screen "Screen_5" 800x480, template "Keep_1"
   Circle "Circle_2" at 38,164 size 32x32
      Appearance <- "Barcode181"
   Circle "Circle_1" at 38,224 size 32x32
      Appearance <- "Barcode190"
   Circle "Circle_3" at 38,279 size 32x32
      Appearance <- "Barcode199"
   Circle "Circle_4" at 38,336 size 32x32
      Appearance <- "Barcode208"
   Circle "Circle_5" at 38,393 size 32x32
      Appearance <- "Barcode217"
   Circle "Circle_6" at 102,164 size 32x32
      Appearance <- "Barcode182"
   Circle "Circle_7" at 102,224 size 32x32
      Appearance <- "Barcode191"
   Circle "Circle_8" at 102,279 size 32x32
      Appearance <- "Barcode200"
   Circle "Circle_9" at 102,336 size 32x32
      Appearance <- "Barcode209"
   Circle "Circle_10" at 102,393 size 32x32
      Appearance <- "Barcode218"
   Circle "Circle_11" at 166,164 size 32x32
      Appearance <- "Barcode183"
   Circle "Circle_12" at 166,224 size 32x32
      Appearance <- "Barcode192"
   Circle "Circle_13" at 166,279 size 32x32
      Appearance <- "Barcode201"
   Circle "Circle_14" at 166,336 size 32x32
      Appearance <- "Barcode210"
   Circle "Circle_15" at 166,393 size 32x32
      Appearance <- "Barcode219"
   Circle "Circle_16" at 230,164 size 32x32
      Appearance <- "Barcode184"
   Circle "Circle_17" at 230,224 size 32x32
      Appearance <- "Barcode193"
   Circle "Circle_18" at 230,279 size 32x32
      Appearance <- "Barcode202"
   Circle "Circle_19" at 230,336 size 32x32
      Appearance <- "Barcode211"
   Circle "Circle_20" at 230,393 size 32x32
      Appearance <- "Barcode220"
   Circle "Circle_21" at 294,164 size 32x32
      Appearance <- "Barcode185"
   Circle "Circle_22" at 294,224 size 32x32
      Appearance <- "Barcode194"
   Circle "Circle_23" at 294,279 size 32x32
      Appearance <- "Barcode203"
   Circle "Circle_24" at 294,336 size 32x32
      Appearance <- "Barcode212"
   Circle "Circle_25" at 294,393 size 32x32
      Appearance <- "Barcode221"
   Circle "Circle_26" at 358,164 size 32x32
      Appearance <- "Barcode186"
   Circle "Circle_27" at 358,225 size 32x32
      Appearance <- "Barcode195"
   Circle "Circle_28" at 358,279 size 32x32
      Appearance <- "Barcode204"
   Circle "Circle_29" at 358,336 size 32x32
      Appearance <- "Barcode213"
   Circle "Circle_30" at 358,393 size 32x32
      Appearance <- "Barcode222"
   Circle "Circle_31" at 422,164 size 32x32
      Appearance <- "Barcode187"
   Circle "Circle_32" at 422,224 size 32x32
      Appearance <- "Barcode196"
   Circle "Circle_33" at 422,279 size 32x32
      Appearance <- "Barcode205"
   Circle "Circle_34" at 422,336 size 32x32
      Appearance <- "Barcode214"
   Circle "Circle_35" at 422,393 size 32x32
      Appearance <- "Barcode223"
   Circle "Circle_36" at 486,164 size 32x32
      Appearance <- "Barcode188"
   Circle "Circle_37" at 486,224 size 32x32
      Appearance <- "Barcode197"
   Circle "Circle_38" at 486,279 size 32x32
      Appearance <- "Barcode206"
   Circle "Circle_39" at 486,336 size 32x32
      Appearance <- "Barcode215"
   Circle "Circle_40" at 486,393 size 32x32
      Appearance <- "Barcode224"
   Circle "Circle_41" at 550,163 size 32x32
      Appearance <- "Barcode189"
   Circle "Circle_42" at 550,224 size 32x32
      Appearance <- "Barcode198"
   Circle "Circle_43" at 550,279 size 32x32
      Appearance <- "Barcode207"
   Circle "Circle_44" at 550,336 size 32x32
      Appearance <- "Barcode216"
   Circle "Circle_45" at 550,393 size 32x32
      Appearance <- "Barcode225"
   TextField "Text field_8" at 473,145 size 66x20; Text 'Box_188'
   TextField "Text field_10" at 25,206 size 66x20; Text 'Box_190'
   TextField "Text field_11" at 88,206 size 66x20; Text 'Box_191'
   TextField "Text field_12" at 153,206 size 66x20; Text 'Box_192'
   TextField "Text field_13" at 217,206 size 66x20; Text 'Box_193'
   TextField "Text field_14" at 281,206 size 66x20; Text 'Box_194'
   TextField "Text field_15" at 345,206 size 66x20; Text 'Box_195'
   TextField "Text field_16" at 410,206 size 66x20; Text 'Box_196'
   TextField "Text field_17" at 473,206 size 66x20; Text 'Box_197'
   TextField "Text field_19" at 26,261 size 66x20; Text 'Box_199'
   TextField "Text field_20" at 89,261 size 66x20; Text 'Box_200'
   TextField "Text field_21" at 153,261 size 66x20; Text 'Box_201'
   TextField "Text field_22" at 217,261 size 66x20; Text 'Box_202'
   TextField "Text field_23" at 281,261 size 66x20; Text 'Box_203'
   TextField "Text field_24" at 346,261 size 66x20; Text 'Box_204'
   TextField "Text field_25" at 409,261 size 66x20; Text 'Box_205'
   TextField "Text field_26" at 473,261 size 66x20; Text 'Box_206'
   TextField "Text field_28" at 25,317 size 66x20; Text 'Box_208'
   TextField "Text field_29" at 88,317 size 66x20; Text 'Box_209'
   TextField "Text field_30" at 153,317 size 66x20; Text 'Box_210'
   TextField "Text field_31" at 218,317 size 66x20; Text 'Box_211'
   TextField "Text field_32" at 282,317 size 66x20; Text 'Box_212'
   TextField "Text field_33" at 346,317 size 66x20; Text 'Box_213'
   TextField "Text field_34" at 410,317 size 66x20; Text 'Box_214'
   TextField "Text field_35" at 472,317 size 66x20; Text 'Box_215'
   TextField "Text field_37" at 26,375 size 66x20; Text 'Box_217'
   TextField "Text field_38" at 88,375 size 66x20; Text 'Box_218'
   TextField "Text field_39" at 153,375 size 66x20; Text 'Box_219'
   TextField "Text field_40" at 217,375 size 66x20; Text 'Box_220'
   TextField "Text field_41" at 281,375 size 66x20; Text 'Box_221'
   TextField "Text field_42" at 345,375 size 66x20; Text 'Box_222'
   TextField "Text field_43" at 409,375 size 66x20; Text 'Box_223'
   TextField "Text field_44" at 473,375 size 66x20; Text 'Box_224'
   TextField "Text field_1" at 24,145 size 66x20; Text 'Box_181'
   TextField "Text field_2" at 87,145 size 66x20; Text 'Box_182'
   TextField "Text field_3" at 152,145 size 66x20; Text 'Box_183'
   TextField "Text field_4" at 216,145 size 66x20; Text 'Box_184'
   TextField "Text field_5" at 280,145 size 66x20; Text 'Box_185'
   TextField "Text field_6" at 344,145 size 66x20; Text 'Box_186'
   TextField "Text field_7" at 409,145 size 66x20; Text 'Box_187'
   TextField "Text field_9" at 536,145 size 66x20; Text 'Box_189'
   TextField "Text field_18" at 537,206 size 66x20; Text 'Box_198'
   TextField "Text field_27" at 537,261 size 66x20; Text 'Box_207'
   TextField "Text field_36" at 537,317 size 66x20; Text 'Box_216'
   TextField "Text field_45" at 536,375 size 66x20; Text 'Box_225'
   SymbolicIOField "Symbolic I/O field_1" at 621,342 size 167x24; TextOn '1'; TextOff '0'; TextList "BOX_All"
      ProcessValue <- "แสดงชื่อยา2"
   IOField "I/O field_1" at 624,160 size 160x64; FormatPattern ???????????
      on OnFinishInput: "Test2"(); "Storage"()
      ProcessValue <- "Expected/Value_All_V"
   TextField "Text field_47" at 648,418 size 78x17; Text ': Low Stock'
   TextField "Text field_46" at 646,395 size 104x17; Text ': Medium Stock'
   TextField "Text field_48" at 646,372 size 82x17; Text ': High Stock'
   GraphicView "Template_Graphic view_6" at 16,8 size 70x68; Picture "KMUTNB-Photoroom"
   GraphicView "Template_Graphic view_5" at 657,59 size 104x124; Picture "channels4_profile-Photoroom"
   Button "Button_5" at 633,292 size 64x24; TextOff 'Back'
      on Click: ActivateScreen("Screen_4", 0)
   Button "Button_6" at 716,292 size 64x24; TextOff 'Next'
      on Click: ActivateScreen("Screen_6", 0)
   GraphicView "Template_Graphic view_1" at 736,255 size 28x26; Picture "NEW_HOME"
   GraphicView "Template_Graphic view_2" at 650,253 size 28x27; Picture "play"
   GraphicView "Template_Graphic view_3" at 721,296 size 20x17; Picture "next-track"
   GraphicView "Template_Graphic view_4" at 638,296 size 20x17; Picture "previous-track"
   Button "Button_3" at 707,246 size 80x42; TextOn 'LOGOUT'; TextOff 'Text'
      on Activate: function_f23ef4c9(); ActivateScreen("1_OVERVIEW_1", 0)
   Button "Button_1" at 623,245 size 80x42; TextOff 'Text'
      on Press: SetTag("มีการปุ่มกดยืนยัน", 1)
      on Release: SetTag("มีการปุ่มกดยืนยัน", 0)
      on Activate: "Storage"()
      on Click: "Conveyor"(); ActivateScreen("Status System", 0)
   TextField "Text field_49" at 734,229 size 32x14; Text 'HOME'
   TextField "Text field_50" at 625,229 size 95x16; Text 'Simmulation Conveyor'

screen "Screen_6" 800x480, template "Keep_1"
   Circle "Circle_2" at 38,164 size 32x32
      Appearance <- "Barcode226"
   Circle "Circle_1" at 38,224 size 32x32
      Appearance <- "Barcode235"
   Circle "Circle_3" at 38,279 size 32x32
      Appearance <- "Barcode244"
   Circle "Circle_4" at 38,336 size 32x32
      Appearance <- "Barcode253"
   Circle "Circle_5" at 38,393 size 32x32
      Appearance <- "Barcode262"
   Circle "Circle_6" at 102,164 size 32x32
      Appearance <- "Barcode227"
   Circle "Circle_7" at 102,224 size 32x32
      Appearance <- "Barcode236"
   Circle "Circle_8" at 102,279 size 32x32
      Appearance <- "Barcode245"
   Circle "Circle_9" at 102,336 size 32x32
      Appearance <- "Barcode254"
   Circle "Circle_10" at 102,393 size 32x32
      Appearance <- "Barcode263"
   Circle "Circle_11" at 166,164 size 32x32
      Appearance <- "Barcode228"
   Circle "Circle_12" at 166,224 size 32x32
      Appearance <- "Barcode237"
   Circle "Circle_13" at 166,279 size 32x32
      Appearance <- "Barcode246"
   Circle "Circle_14" at 166,336 size 32x32
      Appearance <- "Barcode255"
   Circle "Circle_15" at 166,393 size 32x32
      Appearance <- "Barcode264"
   Circle "Circle_16" at 230,164 size 32x32
      Appearance <- "Barcode229"
   Circle "Circle_17" at 230,224 size 32x32
      Appearance <- "Barcode238"
   Circle "Circle_18" at 230,279 size 32x32
      Appearance <- "Barcode247"
   Circle "Circle_19" at 230,336 size 32x32
      Appearance <- "Barcode256"
   Circle "Circle_20" at 230,393 size 32x32
      Appearance <- "Barcode265"
   Circle "Circle_21" at 294,164 size 32x32
      Appearance <- "Barcode230"
   Circle "Circle_22" at 294,224 size 32x32
      Appearance <- "Barcode239"
   Circle "Circle_23" at 294,279 size 32x32
      Appearance <- "Barcode248"
   Circle "Circle_24" at 294,336 size 32x32
      Appearance <- "Barcode257"
   Circle "Circle_25" at 294,393 size 32x32
      Appearance <- "Barcode266"
   Circle "Circle_26" at 358,164 size 32x32
      Appearance <- "Barcode231"
   Circle "Circle_27" at 358,225 size 32x32
      Appearance <- "Barcode240"
   Circle "Circle_28" at 358,279 size 32x32
      Appearance <- "Barcode249"
   Circle "Circle_29" at 358,336 size 32x32
      Appearance <- "Barcode258"
   Circle "Circle_30" at 358,393 size 32x32
      Appearance <- "Barcode267"
   Circle "Circle_31" at 422,164 size 32x32
      Appearance <- "Barcode232"
   Circle "Circle_32" at 422,224 size 32x32
      Appearance <- "Barcode241"
   Circle "Circle_33" at 422,279 size 32x32
      Appearance <- "Barcode250"
   Circle "Circle_34" at 422,336 size 32x32
      Appearance <- "Barcode259"
   Circle "Circle_35" at 422,393 size 32x32
      Appearance <- "Barcode268"
   Circle "Circle_36" at 486,164 size 32x32
      Appearance <- "Barcode233"
   Circle "Circle_37" at 486,224 size 32x32
      Appearance <- "Barcode242"
   Circle "Circle_38" at 486,279 size 32x32
      Appearance <- "Barcode251"
   Circle "Circle_39" at 486,336 size 32x32
      Appearance <- "Barcode260"
   Circle "Circle_40" at 486,393 size 32x32
      Appearance <- "Barcode269"
   Circle "Circle_41" at 550,163 size 32x32
      Appearance <- "Barcode234"
   Circle "Circle_42" at 550,224 size 32x32
      Appearance <- "Barcode243"
   Circle "Circle_43" at 550,279 size 32x32
      Appearance <- "Barcode252"
   Circle "Circle_44" at 550,336 size 32x32
      Appearance <- "Barcode261"
   Circle "Circle_45" at 550,393 size 32x32
      Appearance <- "Barcode270"
   TextField "Text field_8" at 473,145 size 66x20; Text 'Box_233'
   TextField "Text field_10" at 25,206 size 66x20; Text 'Box_235'
   TextField "Text field_11" at 88,206 size 66x20; Text 'Box_236'
   TextField "Text field_12" at 153,206 size 66x20; Text 'Box_237'
   TextField "Text field_13" at 217,206 size 66x20; Text 'Box_238'
   TextField "Text field_14" at 281,206 size 66x20; Text 'Box_239'
   TextField "Text field_15" at 345,206 size 66x20; Text 'Box_240'
   TextField "Text field_16" at 410,206 size 66x20; Text 'Box_241'
   TextField "Text field_17" at 473,206 size 66x20; Text 'Box_242'
   TextField "Text field_19" at 26,261 size 66x20; Text 'Box_244'
   TextField "Text field_20" at 89,261 size 66x20; Text 'Box_245'
   TextField "Text field_21" at 153,261 size 66x20; Text 'Box_246'
   TextField "Text field_22" at 217,261 size 66x20; Text 'Box_247'
   TextField "Text field_23" at 281,261 size 66x20; Text 'Box_248'
   TextField "Text field_24" at 346,261 size 66x20; Text 'Box_249'
   TextField "Text field_25" at 409,261 size 66x20; Text 'Box_250'
   TextField "Text field_26" at 473,261 size 66x20; Text 'Box_251'
   TextField "Text field_28" at 25,317 size 66x20; Text 'Box_253'
   TextField "Text field_29" at 88,317 size 66x20; Text 'Box_254'
   TextField "Text field_30" at 153,317 size 66x20; Text 'Box_255'
   TextField "Text field_31" at 217,317 size 66x20; Text 'Box_256'
   TextField "Text field_32" at 281,317 size 66x20; Text 'Box_257'
   TextField "Text field_33" at 344,317 size 66x20; Text 'Box_258'
   TextField "Text field_34" at 409,317 size 66x20; Text 'Box_259'
   TextField "Text field_35" at 472,317 size 66x20; Text 'Box_260'
   TextField "Text field_37" at 24,375 size 66x20; Text 'Box_262'
   TextField "Text field_38" at 88,375 size 66x20; Text 'Box_263'
   TextField "Text field_39" at 153,375 size 66x20; Text 'Box_264'
   TextField "Text field_40" at 217,375 size 66x20; Text 'Box_265'
   TextField "Text field_41" at 281,375 size 66x20; Text 'Box_266'
   TextField "Text field_42" at 345,375 size 66x20; Text 'Box_267'
   TextField "Text field_43" at 409,375 size 66x20; Text 'Box_268'
   TextField "Text field_44" at 473,375 size 66x20; Text 'Box_269'
   TextField "Text field_1" at 24,145 size 66x20; Text 'Box_226'
   TextField "Text field_2" at 87,145 size 66x20; Text 'Box_227'
   TextField "Text field_3" at 152,145 size 66x20; Text 'Box_228'
   TextField "Text field_4" at 216,145 size 66x20; Text 'Box_229'
   TextField "Text field_5" at 280,145 size 66x20; Text 'Box_230'
   TextField "Text field_6" at 344,145 size 66x20; Text 'Box_231'
   TextField "Text field_7" at 409,145 size 66x20; Text 'Box_232'
   TextField "Text field_9" at 536,145 size 66x20; Text 'Box_234'
   TextField "Text field_18" at 537,206 size 66x20; Text 'Box_243'
   TextField "Text field_27" at 537,261 size 66x20; Text 'Box_252'
   TextField "Text field_36" at 537,317 size 66x20; Text 'Box_261'
   TextField "Text field_45" at 536,375 size 66x20; Text 'Box_270'
   SymbolicIOField "Symbolic I/O field_1" at 621,342 size 167x24; TextOn '1'; TextOff '0'; TextList "BOX_All"
      ProcessValue <- "แสดงชื่อยา2"
   IOField "I/O field_1" at 624,160 size 160x64; FormatPattern ???????????
      on OnFinishInput: "Test2"(); "Storage"()
      ProcessValue <- "Expected/Value_All_V"
   TextField "Text field_47" at 648,418 size 78x17; Text ': Low Stock'
   TextField "Text field_46" at 646,395 size 104x17; Text ': Medium Stock'
   TextField "Text field_48" at 646,372 size 82x17; Text ': High Stock'
   GraphicView "Template_Graphic view_6" at 16,8 size 70x68; Picture "KMUTNB-Photoroom"
   GraphicView "Template_Graphic view_5" at 657,59 size 104x124; Picture "channels4_profile-Photoroom"
   Button "Button_5" at 633,292 size 64x24; TextOff 'Back'
      on Click: ActivateScreen("Screen_5", 0)
   Button "Button_6" at 716,292 size 64x24; TextOff 'Next'
      on Click: ActivateScreen("Screen_7", 0)
   GraphicView "Template_Graphic view_1" at 736,255 size 28x26; Picture "NEW_HOME"
   GraphicView "Template_Graphic view_2" at 650,253 size 28x27; Picture "play"
   GraphicView "Template_Graphic view_3" at 721,296 size 20x17; Picture "next-track"
   GraphicView "Template_Graphic view_4" at 638,296 size 20x17; Picture "previous-track"
   Button "Button_3" at 707,246 size 80x42; TextOn 'LOGOUT'; TextOff 'Text'
      on Activate: function_f23ef4c9(); ActivateScreen("1_OVERVIEW_1", 0)
   Button "Button_1" at 623,245 size 80x42; TextOff 'Text'
      on Press: SetTag("มีการปุ่มกดยืนยัน", 1)
      on Release: SetTag("มีการปุ่มกดยืนยัน", 0)
      on Activate: "Storage"()
      on Click: "Conveyor"(); ActivateScreen("Status System", 0)
   TextField "Text field_49" at 734,229 size 32x14; Text 'HOME'
   TextField "Text field_50" at 625,229 size 95x16; Text 'Simmulation Conveyor'

screen "Screen_7" 800x480, template "Keep_1"
   Circle "Circle_2" at 38,164 size 32x32
      Appearance <- "Barcode271"
   Circle "Circle_1" at 38,224 size 32x32
      Appearance <- "Barcode280"
   Circle "Circle_3" at 38,279 size 32x32
      Appearance <- "Barcode289"
   Circle "Circle_4" at 38,336 size 32x32
      Appearance <- "Barcode298"
   Circle "Circle_5" at 38,393 size 32x32
      Appearance <- "Barcode307"
   Circle "Circle_6" at 102,164 size 32x32
      Appearance <- "Barcode272"
   Circle "Circle_7" at 102,224 size 32x32
      Appearance <- "Barcode281"
   Circle "Circle_8" at 102,279 size 32x32
      Appearance <- "Barcode290"
   Circle "Circle_9" at 102,336 size 32x32
      Appearance <- "Barcode299"
   Circle "Circle_10" at 102,393 size 32x32
      Appearance <- "Barcode308"
   Circle "Circle_11" at 166,164 size 32x32
      Appearance <- "Barcode273"
   Circle "Circle_12" at 166,224 size 32x32
      Appearance <- "Barcode282"
   Circle "Circle_13" at 166,279 size 32x32
      Appearance <- "Barcode291"
   Circle "Circle_14" at 166,336 size 32x32
      Appearance <- "Barcode300"
   Circle "Circle_15" at 166,393 size 32x32
      Appearance <- "Barcode309"
   Circle "Circle_16" at 230,164 size 32x32
      Appearance <- "Barcode274"
   Circle "Circle_17" at 230,224 size 32x32
      Appearance <- "Barcode283"
   Circle "Circle_18" at 230,279 size 32x32
      Appearance <- "Barcode292"
   Circle "Circle_19" at 230,336 size 32x32
      Appearance <- "Barcode301"
   Circle "Circle_20" at 230,393 size 32x32
      Appearance <- "Barcode310"
   Circle "Circle_21" at 294,164 size 32x32
      Appearance <- "Barcode275"
   Circle "Circle_22" at 294,224 size 32x32
      Appearance <- "Barcode284"
   Circle "Circle_23" at 294,279 size 32x32
      Appearance <- "Barcode293"
   Circle "Circle_24" at 294,336 size 32x32
      Appearance <- "Barcode302"
   Circle "Circle_25" at 294,393 size 32x32
      Appearance <- "Barcode311"
   Circle "Circle_26" at 358,164 size 32x32
      Appearance <- "Barcode276"
   Circle "Circle_27" at 358,225 size 32x32
      Appearance <- "Barcode285"
   Circle "Circle_28" at 358,279 size 32x32
      Appearance <- "Barcode294"
   Circle "Circle_29" at 358,336 size 32x32
      Appearance <- "Barcode303"
   Circle "Circle_30" at 358,393 size 32x32
      Appearance <- "Barcode312"
   Circle "Circle_31" at 422,164 size 32x32
      Appearance <- "Barcode277"
   Circle "Circle_32" at 422,224 size 32x32
      Appearance <- "Barcode286"
   Circle "Circle_33" at 422,279 size 32x32
      Appearance <- "Barcode295"
   Circle "Circle_34" at 422,336 size 32x32
      Appearance <- "Barcode304"
   Circle "Circle_35" at 422,393 size 32x32
      Appearance <- "Barcode313"
   Circle "Circle_36" at 486,164 size 32x32
      Appearance <- "Barcode278"
   Circle "Circle_37" at 486,224 size 32x32
      Appearance <- "Barcode287"
   Circle "Circle_38" at 486,279 size 32x32
      Appearance <- "Barcode296"
   Circle "Circle_39" at 486,336 size 32x32
      Appearance <- "Barcode305"
   Circle "Circle_40" at 486,393 size 32x32
      Appearance <- "Barcode314"
   Circle "Circle_41" at 550,163 size 32x32
      Appearance <- "Barcode279"
   Circle "Circle_42" at 550,224 size 32x32
      Appearance <- "Barcode288"
   Circle "Circle_43" at 550,279 size 32x32
      Appearance <- "Barcode297"
   Circle "Circle_44" at 550,336 size 32x32
      Appearance <- "Barcode306"
   Circle "Circle_45" at 550,393 size 32x32
      Appearance <- "Barcode315"
   TextField "Text field_8" at 473,145 size 66x20; Text 'Box_278'
   TextField "Text field_10" at 25,206 size 66x20; Text 'Box_280'
   TextField "Text field_11" at 88,206 size 66x20; Text 'Box_281'
   TextField "Text field_12" at 153,206 size 66x20; Text 'Box_282'
   TextField "Text field_13" at 217,206 size 66x20; Text 'Box_283'
   TextField "Text field_14" at 281,206 size 66x20; Text 'Box_284'
   TextField "Text field_15" at 345,206 size 66x20; Text 'Box_285'
   TextField "Text field_16" at 410,206 size 66x20; Text 'Box_286'
   TextField "Text field_17" at 473,206 size 66x20; Text 'Box_287'
   TextField "Text field_19" at 25,261 size 66x20; Text 'Box_289'
   TextField "Text field_20" at 89,261 size 66x20; Text 'Box_290'
   TextField "Text field_21" at 153,261 size 66x20; Text 'Box_291'
   TextField "Text field_22" at 217,261 size 66x20; Text 'Box_292'
   TextField "Text field_23" at 281,261 size 66x20; Text 'Box_293'
   TextField "Text field_24" at 346,261 size 66x20; Text 'Box_294'
   TextField "Text field_25" at 409,261 size 66x20; Text 'Box_295'
   TextField "Text field_26" at 473,261 size 66x20; Text 'Box_296'
   TextField "Text field_28" at 25,317 size 66x20; Text 'Box_298'
   TextField "Text field_29" at 88,317 size 66x20; Text 'Box_299'
   TextField "Text field_30" at 153,317 size 66x20; Text 'Box_300'
   TextField "Text field_31" at 217,317 size 66x20; Text 'Box_301'
   TextField "Text field_32" at 281,317 size 66x20; Text 'Box_302'
   TextField "Text field_33" at 344,317 size 66x20; Text 'Box_303'
   TextField "Text field_34" at 409,317 size 66x20; Text 'Box_304'
   TextField "Text field_35" at 472,317 size 66x20; Text 'Box_305'
   TextField "Text field_37" at 24,375 size 66x20; Text 'Box_307'
   TextField "Text field_38" at 88,375 size 66x20; Text 'Box_308'
   TextField "Text field_39" at 153,375 size 66x20; Text 'Box_309'
   TextField "Text field_40" at 217,375 size 66x20; Text 'Box_310'
   TextField "Text field_41" at 281,375 size 66x20; Text 'Box_311'
   TextField "Text field_42" at 345,375 size 66x20; Text 'Box_312'
   TextField "Text field_43" at 409,375 size 66x20; Text 'Box_313'
   TextField "Text field_44" at 473,375 size 66x20; Text 'Box_314'
   TextField "Text field_1" at 24,145 size 66x20; Text 'Box_271'
   TextField "Text field_2" at 87,145 size 66x20; Text 'Box_272'
   TextField "Text field_3" at 152,145 size 66x20; Text 'Box_273'
   TextField "Text field_4" at 216,145 size 66x20; Text 'Box_274'
   TextField "Text field_5" at 280,145 size 66x20; Text 'Box_275'
   TextField "Text field_6" at 344,145 size 66x20; Text 'Box_276'
   TextField "Text field_7" at 409,145 size 66x20; Text 'Box_277'
   TextField "Text field_9" at 536,145 size 66x20; Text 'Box_279'
   TextField "Text field_18" at 537,206 size 66x20; Text 'Box_288'
   TextField "Text field_27" at 537,261 size 66x20; Text 'Box_297'
   TextField "Text field_36" at 537,317 size 66x20; Text 'Box_306'
   TextField "Text field_45" at 536,375 size 66x20; Text 'Box_315'
   SymbolicIOField "Symbolic I/O field_1" at 621,342 size 167x24; TextOn '1'; TextOff '0'; TextList "BOX_All"
      ProcessValue <- "แสดงชื่อยา2"
   IOField "I/O field_1" at 624,160 size 160x64; FormatPattern ???????????
      on OnFinishInput: "Test2"(); "Storage"()
      ProcessValue <- "Expected/Value_All_V"
   TextField "Text field_47" at 648,418 size 78x17; Text ': Low Stock'
   TextField "Text field_46" at 646,395 size 104x17; Text ': Medium Stock'
   TextField "Text field_48" at 646,372 size 82x17; Text ': High Stock'
   GraphicView "Template_Graphic view_6" at 16,8 size 70x68; Picture "KMUTNB-Photoroom"
   GraphicView "Template_Graphic view_5" at 657,59 size 104x124; Picture "channels4_profile-Photoroom"
   Button "Button_5" at 633,292 size 64x24; TextOff 'Back'
      on Click: ActivateScreen("Screen_6", 0)
   Button "Button_6" at 716,292 size 64x24; TextOff 'Next'
      on Click: ActivateScreen("Screen_8", 0)
   GraphicView "Template_Graphic view_1" at 736,255 size 28x26; Picture "NEW_HOME"
   GraphicView "Template_Graphic view_2" at 650,253 size 28x27; Picture "play"
   GraphicView "Template_Graphic view_3" at 721,296 size 20x17; Picture "next-track"
   GraphicView "Template_Graphic view_4" at 638,296 size 20x17; Picture "previous-track"
   Button "Button_3" at 707,246 size 80x42; TextOn 'LOGOUT'; TextOff 'Text'
      on Activate: function_f23ef4c9(); ActivateScreen("1_OVERVIEW_1", 0)
   Button "Button_1" at 623,245 size 80x42; TextOff 'Text'
      on Press: SetTag("มีการปุ่มกดยืนยัน", 1)
      on Release: SetTag("มีการปุ่มกดยืนยัน", 0)
      on Activate: "Storage"()
      on Click: "Conveyor"(); ActivateScreen("Status System", 0)
   TextField "Text field_49" at 734,229 size 32x14; Text 'HOME'
   TextField "Text field_50" at 625,229 size 95x16; Text 'Simmulation Conveyor'

screen "Screen_8" 800x480, template "Keep_1"
   Circle "Circle_2" at 38,164 size 32x32
      Appearance <- "Barcode316"
   Circle "Circle_1" at 38,224 size 32x32
      Appearance <- "Barcode325"
   Circle "Circle_3" at 38,279 size 32x32
      Appearance <- "Barcode334"
   Circle "Circle_4" at 38,336 size 32x32
      Appearance <- "Barcode343"
   Circle "Circle_5" at 38,393 size 32x32
      Appearance <- "Barcode352"
   Circle "Circle_6" at 102,164 size 32x32
      Appearance <- "Barcode317"
   Circle "Circle_7" at 102,224 size 32x32
      Appearance <- "Barcode326"
   Circle "Circle_8" at 102,279 size 32x32
      Appearance <- "Barcode335"
   Circle "Circle_9" at 102,336 size 32x32
      Appearance <- "Barcode344"
   Circle "Circle_10" at 102,393 size 32x32
      Appearance <- "Barcode353"
   Circle "Circle_11" at 166,164 size 32x32
      Appearance <- "Barcode318"
   Circle "Circle_12" at 166,224 size 32x32
      Appearance <- "Barcode327"
   Circle "Circle_13" at 166,279 size 32x32
      Appearance <- "Barcode336"
   Circle "Circle_14" at 166,336 size 32x32
      Appearance <- "Barcode345"
   Circle "Circle_15" at 166,393 size 32x32
      Appearance <- "Barcode354"
   Circle "Circle_16" at 230,164 size 32x32
      Appearance <- "Barcode319"
   Circle "Circle_17" at 230,224 size 32x32
      Appearance <- "Barcode328"
   Circle "Circle_18" at 230,279 size 32x32
      Appearance <- "Barcode337"
   Circle "Circle_19" at 230,336 size 32x32
      Appearance <- "Barcode346"
   Circle "Circle_20" at 230,393 size 32x32
      Appearance <- "Barcode355"
   Circle "Circle_21" at 294,164 size 32x32
      Appearance <- "Barcode320"
   Circle "Circle_22" at 294,224 size 32x32
      Appearance <- "Barcode329"
   Circle "Circle_23" at 294,279 size 32x32
      Appearance <- "Barcode338"
   Circle "Circle_24" at 294,336 size 32x32
      Appearance <- "Barcode347"
   Circle "Circle_25" at 294,393 size 32x32
      Appearance <- "Barcode356"
   Circle "Circle_26" at 358,164 size 32x32
      Appearance <- "Barcode321"
   Circle "Circle_27" at 358,225 size 32x32
      Appearance <- "Barcode330"
   Circle "Circle_28" at 358,279 size 32x32
      Appearance <- "Barcode339"
   Circle "Circle_29" at 358,336 size 32x32
      Appearance <- "Barcode348"
   Circle "Circle_30" at 358,393 size 32x32
      Appearance <- "Barcode357"
   Circle "Circle_31" at 422,164 size 32x32
      Appearance <- "Barcode322"
   Circle "Circle_32" at 422,224 size 32x32
      Appearance <- "Barcode331"
   Circle "Circle_33" at 422,279 size 32x32
      Appearance <- "Barcode340"
   Circle "Circle_34" at 422,336 size 32x32
      Appearance <- "Barcode349"
   Circle "Circle_35" at 422,393 size 32x32
      Appearance <- "Barcode358"
   Circle "Circle_36" at 486,164 size 32x32
      Appearance <- "Barcode323"
   Circle "Circle_37" at 486,224 size 32x32
      Appearance <- "Barcode332"
   Circle "Circle_38" at 486,279 size 32x32
      Appearance <- "Barcode341"
   Circle "Circle_39" at 486,336 size 32x32
      Appearance <- "Barcode350"
   Circle "Circle_40" at 486,393 size 32x32
      Appearance <- "Barcode359"
   Circle "Circle_41" at 550,163 size 32x32
      Appearance <- "Barcode324"
   Circle "Circle_42" at 550,224 size 32x32
      Appearance <- "Barcode333"
   Circle "Circle_43" at 550,279 size 32x32
      Appearance <- "Barcode342"
   Circle "Circle_44" at 550,336 size 32x32
      Appearance <- "Barcode351"
   Circle "Circle_45" at 550,393 size 32x32
      Appearance <- "Barcode360"
   TextField "Text field_8" at 473,145 size 66x20; Text 'Box_323'
   TextField "Text field_10" at 25,206 size 66x20; Text 'Box_325'
   TextField "Text field_11" at 88,206 size 66x20; Text 'Box_326'
   TextField "Text field_12" at 153,206 size 66x20; Text 'Box_327'
   TextField "Text field_13" at 217,206 size 66x20; Text 'Box_328'
   TextField "Text field_14" at 281,206 size 66x20; Text 'Box_329'
   TextField "Text field_15" at 345,206 size 66x20; Text 'Box_330'
   TextField "Text field_16" at 410,206 size 66x20; Text 'Box_331'
   TextField "Text field_17" at 473,206 size 66x20; Text 'Box_332'
   TextField "Text field_19" at 25,261 size 66x20; Text 'Box_334'
   TextField "Text field_20" at 89,261 size 66x20; Text 'Box_335'
   TextField "Text field_21" at 153,261 size 66x20; Text 'Box_336'
   TextField "Text field_22" at 217,261 size 66x20; Text 'Box_337'
   TextField "Text field_23" at 281,261 size 66x20; Text 'Box_338'
   TextField "Text field_24" at 346,261 size 66x20; Text 'Box_339'
   TextField "Text field_25" at 409,261 size 66x20; Text 'Box_340'
   TextField "Text field_26" at 473,261 size 66x20; Text 'Box_341'
   TextField "Text field_28" at 25,317 size 66x20; Text 'Box_343'
   TextField "Text field_29" at 88,317 size 66x20; Text 'Box_344'
   TextField "Text field_30" at 153,317 size 66x20; Text 'Box_345'
   TextField "Text field_31" at 217,317 size 66x20; Text 'Box_346'
   TextField "Text field_32" at 281,317 size 66x20; Text 'Box_347'
   TextField "Text field_33" at 344,317 size 66x20; Text 'Box_348'
   TextField "Text field_34" at 409,317 size 66x20; Text 'Box_349'
   TextField "Text field_35" at 472,317 size 66x20; Text 'Box_350'
   TextField "Text field_37" at 24,375 size 66x20; Text 'Box_352'
   TextField "Text field_38" at 88,375 size 66x20; Text 'Box_353'
   TextField "Text field_39" at 153,375 size 66x20; Text 'Box_354'
   TextField "Text field_40" at 217,375 size 66x20; Text 'Box_355'
   TextField "Text field_41" at 281,375 size 66x20; Text 'Box_356'
   TextField "Text field_42" at 345,375 size 66x20; Text 'Box_357'
   TextField "Text field_43" at 409,375 size 66x20; Text 'Box_358'
   TextField "Text field_44" at 473,375 size 66x20; Text 'Box_359'
   TextField "Text field_1" at 24,145 size 66x20; Text 'Box_316'
   TextField "Text field_2" at 89,145 size 66x20; Text 'Box_317'
   TextField "Text field_3" at 152,145 size 66x20; Text 'Box_318'
   TextField "Text field_4" at 216,145 size 66x20; Text 'Box_319'
   TextField "Text field_5" at 280,145 size 66x20; Text 'Box_320'
   TextField "Text field_6" at 344,145 size 66x20; Text 'Box_321'
   TextField "Text field_7" at 409,145 size 66x20; Text 'Box_322'
   TextField "Text field_9" at 536,145 size 66x20; Text 'Box_324'
   TextField "Text field_18" at 537,206 size 66x20; Text 'Box_333'
   TextField "Text field_27" at 537,261 size 66x20; Text 'Box_342'
   TextField "Text field_36" at 537,317 size 66x20; Text 'Box_351'
   TextField "Text field_45" at 536,375 size 66x20; Text 'Box_360'
   SymbolicIOField "Symbolic I/O field_1" at 621,342 size 167x24; TextOn '1'; TextOff '0'; TextList "BOX_All"
      ProcessValue <- "แสดงชื่อยา2"
   IOField "I/O field_1" at 624,160 size 160x64; FormatPattern ???????????
      on OnFinishInput: "Test2"(); "Storage"()
      ProcessValue <- "Expected/Value_All_V"
   TextField "Text field_47" at 648,418 size 78x17; Text ': Low Stock'
   TextField "Text field_46" at 646,395 size 104x17; Text ': Medium Stock'
   TextField "Text field_48" at 646,372 size 82x17; Text ': High Stock'
   GraphicView "Template_Graphic view_6" at 16,8 size 70x68; Picture "KMUTNB-Photoroom"
   GraphicView "Template_Graphic view_5" at 657,59 size 104x124; Picture "channels4_profile-Photoroom"
   Button "Button_5" at 633,292 size 64x24; TextOff 'Back'
      on Click: ActivateScreen("Screen_7", 0)
   Button "Button_6" at 716,292 size 64x24; TextOff 'Next'
      on Click: ActivateScreen("Screen_9", 0)
   GraphicView "Template_Graphic view_1" at 736,255 size 28x26; Picture "NEW_HOME"
   GraphicView "Template_Graphic view_2" at 650,253 size 28x27; Picture "play"
   GraphicView "Template_Graphic view_3" at 721,296 size 20x17; Picture "next-track"
   GraphicView "Template_Graphic view_4" at 638,296 size 20x17; Picture "previous-track"
   Button "Button_3" at 707,246 size 80x42; TextOn 'LOGOUT'; TextOff 'Text'
      on Activate: function_f23ef4c9(); ActivateScreen("1_OVERVIEW_1", 0)
   Button "Button_1" at 623,245 size 80x42; TextOff 'Text'
      on Press: SetTag("มีการปุ่มกดยืนยัน", 1)
      on Release: SetTag("มีการปุ่มกดยืนยัน", 0)
      on Activate: "Storage"()
      on Click: "Conveyor"(); ActivateScreen("Status System", 0)
   TextField "Text field_49" at 734,229 size 32x14; Text 'HOME'
   TextField "Text field_50" at 625,229 size 95x16; Text 'Simmulation Conveyor'

screen "Screen_9" 800x480, template "Keep_1"
   TextField "Text field_8" at 473,145 size 66x20; Text 'Box_368'
   TextField "Text field_10" at 25,206 size 66x20; Text 'Box_370'
   TextField "Text field_11" at 88,206 size 66x20; Text 'Box_371'
   TextField "Text field_12" at 153,206 size 66x20; Text 'Box_372'
   TextField "Text field_13" at 217,206 size 66x20; Text 'Box_373'
   TextField "Text field_14" at 281,206 size 66x20; Text 'Box_374'
   TextField "Text field_15" at 345,206 size 66x20; Text 'Box_375'
   TextField "Text field_16" at 410,206 size 66x20; Text 'Box_376'
   TextField "Text field_17" at 473,206 size 66x20; Text 'Box_377'
   TextField "Text field_19" at 25,261 size 66x20; Text 'Box_379'
   TextField "Text field_20" at 89,261 size 66x20; Text 'Box_380'
   TextField "Text field_21" at 153,261 size 66x20; Text 'Box_381'
   TextField "Text field_22" at 217,261 size 66x20; Text 'Box_382'
   TextField "Text field_23" at 281,261 size 66x20; Text 'Box_383'
   TextField "Text field_24" at 346,261 size 66x20; Text 'Box_384'
   TextField "Text field_25" at 409,261 size 66x20; Text 'Box_385'
   TextField "Text field_26" at 473,261 size 66x20; Text 'Box_386'
   TextField "Text field_28" at 25,317 size 66x20; Text 'Box_388'
   TextField "Text field_29" at 88,317 size 66x20; Text 'Box_389'
   TextField "Text field_30" at 153,317 size 66x20; Text 'Box_390'
   TextField "Text field_31" at 217,317 size 66x20; Text 'Box_391'
   TextField "Text field_32" at 281,317 size 66x20; Text 'Box_392'
   TextField "Text field_33" at 344,317 size 66x20; Text 'Box_393'
   TextField "Text field_34" at 409,317 size 66x20; Text 'Box_394'
   TextField "Text field_35" at 472,317 size 66x20; Text 'Box_395'
   TextField "Text field_37" at 24,375 size 66x20; Text 'Box_397'
   TextField "Text field_38" at 88,375 size 66x20; Text 'Box_398'
   TextField "Text field_39" at 153,375 size 66x20; Text 'Box_399'
   TextField "Text field_40" at 217,375 size 66x20; Text 'Box_400'
   TextField "Text field_41" at 281,375 size 66x20; Text 'Box_401'
   TextField "Text field_42" at 345,375 size 66x20; Text 'Box_402'
   TextField "Text field_43" at 409,375 size 66x20; Text 'Box_403'
   TextField "Text field_44" at 473,375 size 66x20; Text 'Box_404'
   TextField "Text field_1" at 24,145 size 66x20; Text 'Box_361'
   TextField "Text field_2" at 89,145 size 66x20; Text 'Box_362'
   TextField "Text field_3" at 152,145 size 66x20; Text 'Box_363'
   TextField "Text field_4" at 216,145 size 66x20; Text 'Box_364'
   TextField "Text field_5" at 280,145 size 66x20; Text 'Box_365'
   TextField "Text field_6" at 344,145 size 66x20; Text 'Box_366'
   TextField "Text field_7" at 409,145 size 66x20; Text 'Box_367'
   TextField "Text field_9" at 536,145 size 66x20; Text 'Box_369'
   TextField "Text field_18" at 537,206 size 66x20; Text 'Box_378'
   TextField "Text field_27" at 537,261 size 66x20; Text 'Box_387'
   TextField "Text field_36" at 537,317 size 66x20; Text 'Box_396'
   TextField "Text field_45" at 536,375 size 66x20; Text 'Box_405'
   SymbolicIOField "Symbolic I/O field_1" at 621,342 size 167x24; TextOn '1'; TextOff '0'; TextList "BOX_All"
      ProcessValue <- "แสดงชื่อยา2"
   IOField "I/O field_1" at 624,160 size 160x64; FormatPattern ???????????
      on OnFinishInput: "Test2"(); "Storage"()
      ProcessValue <- "Expected/Value_All_V"
   TextField "Text field_47" at 648,418 size 78x17; Text ': Low Stock'
   TextField "Text field_46" at 646,395 size 104x17; Text ': Medium Stock'
   TextField "Text field_48" at 646,372 size 82x17; Text ': High Stock'
   Circle "Circle_2" at 38,164 size 32x32
      Appearance <- "Barcode361"
   Circle "Circle_1" at 38,224 size 32x32
      Appearance <- "Barcode370"
   Circle "Circle_3" at 38,279 size 32x32
      Appearance <- "Barcode379"
   Circle "Circle_4" at 38,336 size 32x32
      Appearance <- "Barcode388"
   Circle "Circle_5" at 38,393 size 32x32
      Appearance <- "Barcode397"
   Circle "Circle_6" at 102,164 size 32x32
      Appearance <- "Barcode362"
   Circle "Circle_7" at 102,224 size 32x32
      Appearance <- "Barcode371"
   Circle "Circle_8" at 102,279 size 32x32
      Appearance <- "Barcode380"
   Circle "Circle_9" at 102,336 size 32x32
      Appearance <- "Barcode389"
   Circle "Circle_10" at 102,393 size 32x32
      Appearance <- "Barcode398"
   Circle "Circle_11" at 166,164 size 32x32
      Appearance <- "Barcode363"
   Circle "Circle_12" at 166,224 size 32x32
      Appearance <- "Barcode372"
   Circle "Circle_13" at 166,279 size 32x32
      Appearance <- "Barcode381"
   Circle "Circle_14" at 166,336 size 32x32
      Appearance <- "Barcode390"
   Circle "Circle_15" at 166,393 size 32x32
      Appearance <- "Barcode399"
   Circle "Circle_16" at 230,164 size 32x32
      Appearance <- "Barcode364"
   Circle "Circle_17" at 230,224 size 32x32
      Appearance <- "Barcode373"
   Circle "Circle_18" at 230,279 size 32x32
      Appearance <- "Barcode382"
   Circle "Circle_19" at 230,336 size 32x32
      Appearance <- "Barcode391"
   Circle "Circle_20" at 230,393 size 32x32
      Appearance <- "Barcode400"
   Circle "Circle_21" at 294,164 size 32x32
      Appearance <- "Barcode365"
   Circle "Circle_22" at 294,224 size 32x32
      Appearance <- "Barcode374"
   Circle "Circle_23" at 294,279 size 32x32
      Appearance <- "Barcode383"
   Circle "Circle_24" at 294,336 size 32x32
      Appearance <- "Barcode392"
   Circle "Circle_25" at 294,393 size 32x32
      Appearance <- "Barcode401"
   Circle "Circle_26" at 358,164 size 32x32
      Appearance <- "Barcode366"
   Circle "Circle_27" at 358,225 size 32x32
      Appearance <- "Barcode375"
   Circle "Circle_28" at 358,279 size 32x32
      Appearance <- "Barcode384"
   Circle "Circle_29" at 358,336 size 32x32
      Appearance <- "Barcode393"
   Circle "Circle_30" at 358,393 size 32x32
      Appearance <- "Barcode402"
   Circle "Circle_31" at 422,164 size 32x32
      Appearance <- "Barcode367"
   Circle "Circle_32" at 422,224 size 32x32
      Appearance <- "Barcode376"
   Circle "Circle_33" at 422,279 size 32x32
      Appearance <- "Barcode385"
   Circle "Circle_34" at 422,336 size 32x32
      Appearance <- "Barcode394"
   Circle "Circle_35" at 422,393 size 32x32
      Appearance <- "Barcode403"
   Circle "Circle_36" at 486,164 size 32x32
      Appearance <- "Barcode368"
   Circle "Circle_37" at 486,224 size 32x32
      Appearance <- "Barcode377"
   Circle "Circle_38" at 486,279 size 32x32
      Appearance <- "Barcode386"
   Circle "Circle_39" at 486,336 size 32x32
      Appearance <- "Barcode395"
   Circle "Circle_40" at 486,393 size 32x32
      Appearance <- "Barcode404"
   Circle "Circle_41" at 550,163 size 32x32
      Appearance <- "Barcode369"
   Circle "Circle_42" at 550,224 size 32x32
      Appearance <- "Barcode378"
   Circle "Circle_43" at 550,279 size 32x32
      Appearance <- "Barcode387"
   Circle "Circle_44" at 550,336 size 32x32
      Appearance <- "Barcode396"
   Circle "Circle_45" at 550,393 size 32x32
      Appearance <- "Barcode405"
   GraphicView "Template_Graphic view_6" at 16,8 size 70x68; Picture "KMUTNB-Photoroom"
   GraphicView "Template_Graphic view_5" at 657,59 size 104x124; Picture "channels4_profile-Photoroom"
   Button "Button_5" at 633,292 size 64x24; TextOff 'Back'
      on Click: ActivateScreen("Screen_8", 0)
   Button "Button_6" at 716,292 size 64x24; TextOff 'Next'
      on Click: ActivateScreen("Screen_10", 0)
   GraphicView "Template_Graphic view_1" at 736,255 size 28x26; Picture "NEW_HOME"
   GraphicView "Template_Graphic view_2" at 650,253 size 28x27; Picture "play"
   GraphicView "Template_Graphic view_3" at 721,296 size 20x17; Picture "next-track"
   GraphicView "Template_Graphic view_4" at 638,296 size 20x17; Picture "previous-track"
   Button "Button_3" at 707,246 size 80x42; TextOn 'LOGOUT'; TextOff 'Text'
      on Activate: function_f23ef4c9(); ActivateScreen("1_OVERVIEW_1", 0)
   Button "Button_1" at 623,245 size 80x42; TextOff 'Text'
      on Press: SetTag("มีการปุ่มกดยืนยัน", 1)
      on Release: SetTag("มีการปุ่มกดยืนยัน", 0)
      on Activate: "Storage"()
      on Click: "Conveyor"(); ActivateScreen("Status System", 0)
   TextField "Text field_49" at 734,229 size 32x14; Text 'HOME'
   TextField "Text field_50" at 625,229 size 95x16; Text 'Simmulation Conveyor'

screen "Screen_10" 800x480, template "Keep_1"
   TextField "Text field_8" at 473,145 size 66x20; Text 'Box_413'
   TextField "Text field_10" at 25,206 size 66x20; Text 'Box_415'
   TextField "Text field_11" at 88,206 size 66x20; Text 'Box_416'
   TextField "Text field_12" at 153,206 size 66x20; Text 'Box_417'
   TextField "Text field_13" at 217,206 size 66x20; Text 'Box_418'
   TextField "Text field_14" at 281,206 size 66x20; Text 'Box_419'
   TextField "Text field_15" at 345,206 size 66x20; Text 'Box_420'
   TextField "Text field_16" at 410,206 size 66x20; Text 'Box_421'
   TextField "Text field_17" at 473,206 size 66x20; Text 'Box_422'
   TextField "Text field_19" at 25,261 size 66x20; Text 'Box_424'
   TextField "Text field_20" at 89,261 size 66x20; Text 'Box_425'
   TextField "Text field_21" at 153,261 size 66x20; Text 'Box_426'
   TextField "Text field_22" at 217,261 size 66x20; Text 'Box_427'
   TextField "Text field_23" at 281,261 size 66x20; Text 'Box_428'
   TextField "Text field_24" at 346,261 size 66x20; Text 'Box_429'
   TextField "Text field_25" at 409,261 size 66x20; Text 'Box_430'
   TextField "Text field_26" at 473,261 size 66x20; Text 'Box_431'
   TextField "Text field_28" at 25,317 size 66x20; Text 'Box_433'
   TextField "Text field_29" at 88,317 size 66x20; Text 'Box_434'
   TextField "Text field_30" at 153,317 size 66x20; Text 'Box_435'
   TextField "Text field_31" at 217,317 size 66x20; Text 'Box_436'
   TextField "Text field_32" at 281,317 size 66x20; Text 'Box_437'
   TextField "Text field_33" at 344,317 size 66x20; Text 'Box_438'
   TextField "Text field_34" at 409,317 size 66x20; Text 'Box_439'
   TextField "Text field_35" at 472,317 size 66x20; Text 'Box_440'
   TextField "Text field_37" at 24,375 size 66x20; Text 'Box_442'
   TextField "Text field_38" at 88,375 size 66x20; Text 'Box_443'
   TextField "Text field_39" at 153,375 size 66x20; Text 'Box_444'
   TextField "Text field_40" at 217,375 size 66x20; Text 'Box_445'
   TextField "Text field_41" at 281,375 size 66x20; Text 'Box_446'
   TextField "Text field_42" at 345,375 size 66x20; Text 'Box_447'
   TextField "Text field_43" at 409,375 size 66x20; Text 'Box_448'
   TextField "Text field_44" at 473,375 size 66x20; Text 'Box_449'
   TextField "Text field_1" at 24,145 size 66x20; Text 'Box_406'
   TextField "Text field_2" at 89,145 size 66x20; Text 'Box_407'
   TextField "Text field_3" at 152,145 size 66x20; Text 'Box_408'
   TextField "Text field_4" at 216,145 size 66x20; Text 'Box_409'
   TextField "Text field_5" at 280,145 size 66x20; Text 'Box_410'
   TextField "Text field_6" at 344,145 size 66x20; Text 'Box_411'
   TextField "Text field_7" at 409,145 size 66x20; Text 'Box_412'
   TextField "Text field_9" at 536,145 size 66x20; Text 'Box_414'
   TextField "Text field_18" at 537,206 size 66x20; Text 'Box_423'
   TextField "Text field_27" at 537,261 size 66x20; Text 'Box_432'
   TextField "Text field_36" at 537,317 size 66x20; Text 'Box_441'
   TextField "Text field_45" at 536,375 size 66x20; Text 'Box_450'
   IOField "I/O field_1" at 624,160 size 160x64; FormatPattern ???????????
      on OnFinishInput: "Test2"(); "Storage"()
      ProcessValue <- "Expected/Value_All_V"
   SymbolicIOField "Symbolic I/O field_1" at 621,342 size 167x24; TextOn '1'; TextOff '0'; TextList "BOX_All"
      ProcessValue <- "แสดงชื่อยา2"
   TextField "Text field_47" at 648,418 size 78x17; Text ': Low Stock'
   TextField "Text field_46" at 646,395 size 104x17; Text ': Medium Stock'
   TextField "Text field_48" at 646,372 size 82x17; Text ': High Stock'
   Circle "Circle_2" at 38,164 size 32x32
      Appearance <- "Barcode406"
   Circle "Circle_1" at 38,224 size 32x32
      Appearance <- "Barcode415"
   Circle "Circle_3" at 38,279 size 32x32
      Appearance <- "Barcode424"
   Circle "Circle_4" at 38,336 size 32x32
      Appearance <- "Barcode433"
   Circle "Circle_5" at 38,393 size 32x32
      Appearance <- "Barcode442"
   Circle "Circle_6" at 102,164 size 32x32
      Appearance <- "Barcode407"
   Circle "Circle_7" at 102,224 size 32x32
      Appearance <- "Barcode416"
   Circle "Circle_8" at 102,279 size 32x32
      Appearance <- "Barcode425"
   Circle "Circle_9" at 102,336 size 32x32
      Appearance <- "Barcode434"
   Circle "Circle_10" at 102,393 size 32x32
      Appearance <- "Barcode443"
   Circle "Circle_11" at 166,164 size 32x32
      Appearance <- "Barcode408"
   Circle "Circle_12" at 166,224 size 32x32
      Appearance <- "Barcode417"
   Circle "Circle_13" at 166,279 size 32x32
      Appearance <- "Barcode426"
   Circle "Circle_14" at 166,336 size 32x32
      Appearance <- "Barcode435"
   Circle "Circle_15" at 166,393 size 32x32
      Appearance <- "Barcode444"
   Circle "Circle_16" at 230,164 size 32x32
      Appearance <- "Barcode409"
   Circle "Circle_17" at 230,224 size 32x32
      Appearance <- "Barcode418"
   Circle "Circle_18" at 230,279 size 32x32
      Appearance <- "Barcode427"
   Circle "Circle_19" at 230,336 size 32x32
      Appearance <- "Barcode436"
   Circle "Circle_20" at 230,393 size 32x32
      Appearance <- "Barcode445"
   Circle "Circle_21" at 294,164 size 32x32
      Appearance <- "Barcode410"
   Circle "Circle_22" at 294,224 size 32x32
      Appearance <- "Barcode419"
   Circle "Circle_23" at 296,280 size 32x32
      Appearance <- "Barcode428"
   Circle "Circle_24" at 294,336 size 32x32
      Appearance <- "Barcode437"
   Circle "Circle_25" at 294,393 size 32x32
      Appearance <- "Barcode446"
   Circle "Circle_26" at 358,164 size 32x32
      Appearance <- "Barcode411"
   Circle "Circle_27" at 358,225 size 32x32
      Appearance <- "Barcode420"
   Circle "Circle_28" at 358,279 size 32x32
      Appearance <- "Barcode429"
   Circle "Circle_29" at 358,336 size 32x32
      Appearance <- "Barcode438"
   Circle "Circle_30" at 358,393 size 32x32
      Appearance <- "Barcode447"
   Circle "Circle_31" at 422,164 size 32x32
      Appearance <- "Barcode412"
   Circle "Circle_32" at 422,224 size 32x32
      Appearance <- "Barcode421"
   Circle "Circle_33" at 422,279 size 32x32
      Appearance <- "Barcode430"
   Circle "Circle_34" at 422,336 size 32x32
      Appearance <- "Barcode439"
   Circle "Circle_35" at 422,393 size 32x32
      Appearance <- "Barcode448"
   Circle "Circle_36" at 486,164 size 32x32
      Appearance <- "Barcode413"
   Circle "Circle_37" at 486,224 size 32x32
      Appearance <- "Barcode422"
   Circle "Circle_38" at 486,279 size 32x32
      Appearance <- "Barcode431"
   Circle "Circle_39" at 486,336 size 32x32
      Appearance <- "Barcode440"
   Circle "Circle_40" at 486,393 size 32x32
      Appearance <- "Barcode449"
   Circle "Circle_41" at 550,163 size 32x32
      Appearance <- "Barcode414"
   Circle "Circle_42" at 550,224 size 32x32
      Appearance <- "Barcode423"
   Circle "Circle_43" at 550,279 size 32x32
      Appearance <- "Barcode432"
   Circle "Circle_44" at 550,336 size 32x32
      Appearance <- "Barcode441"
   Circle "Circle_45" at 550,393 size 32x32
      Appearance <- "Barcode450"
   GraphicView "Template_Graphic view_6" at 16,8 size 70x68; Picture "KMUTNB-Photoroom"
   GraphicView "Template_Graphic view_5" at 657,59 size 104x124; Picture "channels4_profile-Photoroom"
   Button "Button_5" at 633,292 size 64x24; TextOff 'Back'
      on Click: ActivateScreen("Screen_9", 0)
   Button "Button_6" at 716,292 size 64x24; TextOff 'Next'
      on Click: ActivateScreen("Screen_11", 0)
   GraphicView "Template_Graphic view_1" at 736,255 size 28x26; Picture "NEW_HOME"
   GraphicView "Template_Graphic view_2" at 650,253 size 28x27; Picture "play"
   GraphicView "Template_Graphic view_3" at 721,296 size 20x17; Picture "next-track"
   GraphicView "Template_Graphic view_4" at 638,296 size 20x17; Picture "previous-track"
   Button "Button_3" at 707,246 size 80x42; TextOn 'LOGOUT'; TextOff 'Text'
      on Activate: function_f23ef4c9(); ActivateScreen("1_OVERVIEW_1", 0)
   Button "Button_1" at 623,245 size 80x42; TextOff 'Text'
      on Press: SetTag("มีการปุ่มกดยืนยัน", 1)
      on Release: SetTag("มีการปุ่มกดยืนยัน", 0)
      on Activate: "Storage"()
      on Click: "Conveyor"(); ActivateScreen("Status System", 0)
   TextField "Text field_49" at 734,229 size 32x14; Text 'HOME'
   TextField "Text field_50" at 625,229 size 95x16; Text 'Simmulation Conveyor'

screen "Screen_11" 800x480, template "Keep_1"
   Circle "Circle_2" at 38,164 size 32x32
      Appearance <- "Barcode451"
   Circle "Circle_1" at 38,224 size 32x32
      Appearance <- "Barcode460"
   Circle "Circle_3" at 38,279 size 32x32
      Appearance <- "Barcode469"
   Circle "Circle_4" at 38,336 size 32x32
      Appearance <- "Barcode478"
   Circle "Circle_5" at 38,393 size 32x32
      Appearance <- "Barcode487"
   Circle "Circle_6" at 102,164 size 32x32
      Appearance <- "Barcode452"
   Circle "Circle_7" at 102,224 size 32x32
      Appearance <- "Barcode461"
   Circle "Circle_8" at 102,279 size 32x32
      Appearance <- "Barcode470"
   Circle "Circle_9" at 102,336 size 32x32
      Appearance <- "Barcode479"
   Circle "Circle_10" at 102,393 size 32x32
      Appearance <- "Barcode488"
   Circle "Circle_11" at 166,164 size 32x32
      Appearance <- "Barcode453"
   Circle "Circle_12" at 166,224 size 32x32
      Appearance <- "Barcode462"
   Circle "Circle_13" at 166,279 size 32x32
      Appearance <- "Barcode471"
   Circle "Circle_14" at 166,336 size 32x32
      Appearance <- "Barcode480"
   Circle "Circle_15" at 166,393 size 32x32
      Appearance <- "Barcode489"
   Circle "Circle_16" at 230,164 size 32x32
      Appearance <- "Barcode454"
   Circle "Circle_17" at 230,224 size 32x32
      Appearance <- "Barcode463"
   Circle "Circle_18" at 230,279 size 32x32
      Appearance <- "Barcode472"
   Circle "Circle_19" at 230,336 size 32x32
      Appearance <- "Barcode481"
   Circle "Circle_20" at 230,393 size 32x32
      Appearance <- "Barcode490"
   Circle "Circle_21" at 294,164 size 32x32
      Appearance <- "Barcode455"
   Circle "Circle_22" at 294,224 size 32x32
      Appearance <- "Barcode464"
   Circle "Circle_23" at 294,279 size 32x32
      Appearance <- "Barcode473"
   Circle "Circle_24" at 294,336 size 32x32
      Appearance <- "Barcode482"
   Circle "Circle_25" at 294,393 size 32x32
      Appearance <- "Barcode491"
   Circle "Circle_26" at 358,164 size 32x32
      Appearance <- "Barcode456"
   Circle "Circle_27" at 358,225 size 32x32
      Appearance <- "Barcode465"
   Circle "Circle_28" at 358,279 size 32x32
      Appearance <- "Barcode474"
   Circle "Circle_29" at 358,336 size 32x32
      Appearance <- "Barcode483"
   Circle "Circle_30" at 358,393 size 32x32
      Appearance <- "Barcode492"
   Circle "Circle_31" at 422,164 size 32x32
      Appearance <- "Barcode457"
   Circle "Circle_32" at 422,224 size 32x32
      Appearance <- "Barcode466"
   Circle "Circle_33" at 422,279 size 32x32
      Appearance <- "Barcode475"
   Circle "Circle_34" at 424,336 size 32x32
      Appearance <- "Barcode484"
   Circle "Circle_35" at 422,393 size 32x32
      Appearance <- "Barcode493"
   Circle "Circle_36" at 486,164 size 32x32
      Appearance <- "Barcode458"
   Circle "Circle_37" at 486,224 size 32x32
      Appearance <- "Barcode467"
   Circle "Circle_38" at 486,279 size 32x32
      Appearance <- "Barcode476"
   Circle "Circle_39" at 486,336 size 32x32
      Appearance <- "Barcode485"
   Circle "Circle_40" at 486,393 size 32x32
      Appearance <- "Barcode494"
   Circle "Circle_41" at 550,163 size 32x32
      Appearance <- "Barcode459"
   Circle "Circle_42" at 550,224 size 32x32
      Appearance <- "Barcode468"
   Circle "Circle_43" at 550,279 size 32x32
      Appearance <- "Barcode477"
   Circle "Circle_44" at 550,336 size 32x32
      Appearance <- "Barcode486"
   TextField "Text field_8" at 473,145 size 66x20; Text 'Box_458'
   TextField "Text field_10" at 25,206 size 66x20; Text 'Box_460'
   TextField "Text field_11" at 88,206 size 66x20; Text 'Box_461'
   TextField "Text field_12" at 153,206 size 66x20; Text 'Box_462'
   TextField "Text field_13" at 217,206 size 66x20; Text 'Box_463'
   TextField "Text field_14" at 281,206 size 66x20; Text 'Box_464'
   TextField "Text field_15" at 345,206 size 66x20; Text 'Box_465'
   TextField "Text field_16" at 410,206 size 66x20; Text 'Box_466'
   TextField "Text field_17" at 473,206 size 66x20; Text 'Box_467'
   TextField "Text field_19" at 25,261 size 66x20; Text 'Box_469'
   TextField "Text field_20" at 89,261 size 66x20; Text 'Box_470'
   TextField "Text field_21" at 153,261 size 66x20; Text 'Box_471'
   TextField "Text field_22" at 217,261 size 66x20; Text 'Box_472'
   TextField "Text field_23" at 281,261 size 66x20; Text 'Box_473'
   TextField "Text field_24" at 346,261 size 66x20; Text 'Box_474'
   TextField "Text field_25" at 409,261 size 66x20; Text 'Box_475'
   TextField "Text field_26" at 473,261 size 66x20; Text 'Box_476'
   TextField "Text field_28" at 25,317 size 66x20; Text 'Box_478'
   TextField "Text field_29" at 88,317 size 66x20; Text 'Box_479'
   TextField "Text field_30" at 153,317 size 66x20; Text 'Box_480'
   TextField "Text field_31" at 217,317 size 66x20; Text 'Box_481'
   TextField "Text field_32" at 281,317 size 66x20; Text 'Box_482'
   TextField "Text field_33" at 344,317 size 66x20; Text 'Box_483'
   TextField "Text field_34" at 409,317 size 66x20; Text 'Box_484'
   TextField "Text field_35" at 472,317 size 66x20; Text 'Box_485'
   TextField "Text field_37" at 24,375 size 66x20; Text 'Box_487'
   TextField "Text field_38" at 88,375 size 66x20; Text 'Box_488'
   TextField "Text field_39" at 153,375 size 66x20; Text 'Box_489'
   TextField "Text field_40" at 217,375 size 66x20; Text 'Box_490'
   TextField "Text field_41" at 281,375 size 66x20; Text 'Box_491'
   TextField "Text field_42" at 345,375 size 66x20; Text 'Box_492'
   TextField "Text field_43" at 409,375 size 66x20; Text 'Box_493'
   TextField "Text field_44" at 473,375 size 66x20; Text 'Box_494'
   TextField "Text field_1" at 24,145 size 66x20; Text 'Box_451'
   TextField "Text field_2" at 89,145 size 66x20; Text 'Box_452'
   TextField "Text field_3" at 152,145 size 66x20; Text 'Box_453'
   TextField "Text field_4" at 216,145 size 66x20; Text 'Box_454'
   TextField "Text field_5" at 280,145 size 66x20; Text 'Box_455'
   TextField "Text field_6" at 344,145 size 66x20; Text 'Box_456'
   TextField "Text field_7" at 409,145 size 66x20; Text 'Box_457'
   TextField "Text field_9" at 536,145 size 66x20; Text 'Box_459'
   TextField "Text field_18" at 537,206 size 66x20; Text 'Box_468'
   TextField "Text field_27" at 537,261 size 66x20; Text 'Box_477'
   TextField "Text field_36" at 537,317 size 66x20; Text 'Box_486'
   IOField "I/O field_1" at 624,160 size 160x64; FormatPattern ???????????
      on OnFinishInput: "Test2"(); "Storage"()
      ProcessValue <- "Expected/Value_All_V"
   SymbolicIOField "Symbolic I/O field_1" at 621,342 size 167x24; TextOn '1'; TextOff '0'; TextList "BOX_All"
      ProcessValue <- "แสดงชื่อยา2"
   TextField "Text field_47" at 648,418 size 78x17; Text ': Low Stock'
   TextField "Text field_46" at 646,395 size 104x17; Text ': Medium Stock'
   TextField "Text field_48" at 646,372 size 82x17; Text ': High Stock'
   GraphicView "Template_Graphic view_6" at 16,8 size 70x68; Picture "KMUTNB-Photoroom"
   GraphicView "Template_Graphic view_5" at 657,59 size 104x124; Picture "channels4_profile-Photoroom"
   Button "Button_5" at 633,292 size 64x24; TextOff 'Back'
      on Click: ActivateScreen("Screen_10", 0)
   GraphicView "Template_Graphic view_1" at 736,255 size 28x26; Picture "NEW_HOME"
   GraphicView "Template_Graphic view_2" at 650,253 size 28x27; Picture "play"
   GraphicView "Template_Graphic view_4" at 638,296 size 20x17; Picture "previous-track"
   Button "Button_3" at 707,246 size 80x42; TextOn 'LOGOUT'; TextOff 'Text'
      on Activate: function_f23ef4c9(); ActivateScreen("1_OVERVIEW_1", 0)
   Button "Button_1" at 623,245 size 80x42; TextOff 'Text'
      on Press: SetTag("มีการปุ่มกดยืนยัน", 1)
      on Release: SetTag("มีการปุ่มกดยืนยัน", 0)
      on Activate: "Storage"()
      on Click: "Conveyor"(); ActivateScreen("Status System", 0)
   TextField "Text field_49" at 734,229 size 32x14; Text 'HOME'
   TextField "Text field_50" at 625,229 size 95x16; Text 'Simmulation Conveyor'

screen "Screen_12" 800x480, template "Keep_1"
   TextField "Text field_8" at 473,145 size 66x20; Text 'Box_503'
   TextField "Text field_10" at 25,206 size 66x20; Text 'Box_505'
   TextField "Text field_11" at 88,206 size 66x20; Text 'Box_506'
   TextField "Text field_12" at 153,206 size 66x20; Text 'Box_507'
   TextField "Text field_13" at 217,206 size 66x20; Text 'Box_508'
   TextField "Text field_14" at 281,206 size 66x20; Text 'Box_509'
   TextField "Text field_15" at 345,206 size 66x20; Text 'Box_510'
   TextField "Text field_16" at 410,206 size 66x20; Text 'Box_511'
   TextField "Text field_17" at 473,206 size 66x20; Text 'Box_512'
   TextField "Text field_19" at 25,261 size 66x20; Text 'Box_514'
   TextField "Text field_20" at 89,261 size 66x20; Text 'Box_515'
   TextField "Text field_21" at 153,261 size 66x20; Text 'Box_516'
   TextField "Text field_22" at 217,261 size 66x20; Text 'Box_517'
   TextField "Text field_23" at 281,261 size 66x20; Text 'Box_518'
   TextField "Text field_24" at 346,261 size 66x20; Text 'Box_519'
   TextField "Text field_25" at 409,261 size 66x20; Text 'Box_520'
   TextField "Text field_1" at 24,145 size 66x20; Text 'Box_496'
   TextField "Text field_2" at 89,145 size 66x20; Text 'Box_497'
   TextField "Text field_3" at 152,145 size 66x20; Text 'Box_498'
   TextField "Text field_4" at 216,145 size 66x20; Text 'Box_499'
   TextField "Text field_5" at 280,145 size 66x20; Text 'Box_500'
   TextField "Text field_6" at 344,145 size 66x20; Text 'Box_501'
   TextField "Text field_7" at 409,145 size 66x20; Text 'Box_502'
   TextField "Text field_9" at 536,145 size 66x20; Text 'Box_504'
   TextField "Text field_18" at 537,206 size 66x20; Text 'Box_513'
   IOField "I/O field_1" at 624,160 size 160x64; FormatPattern ???????????
      on OnFinishInput: "Test2"()
      ProcessValue <- "Expected/Value_All_V"
   SymbolicIOField "Symbolic I/O field_1" at 621,342 size 167x24; TextOn '1'; TextOff '0'; TextList "BOX_All"
      ProcessValue <- "แสดงชื่อยา2"
   TextField "Text field_47" at 648,418 size 78x17; Text ': Low Stock'
   TextField "Text field_46" at 646,395 size 104x17; Text ': Medium Stock'
   TextField "Text field_48" at 646,372 size 82x17; Text ': High Stock'
   Circle "Circle_2" at 38,164 size 32x32
      Appearance <- "Barcode496"
   Circle "Circle_1" at 38,224 size 32x32
      Appearance <- "Barcode505"
   Circle "Circle_3" at 38,279 size 32x32
      Appearance <- "Barcode514"
   Circle "Circle_6" at 102,164 size 32x32
      Appearance <- "Barcode497"
   Circle "Circle_7" at 102,224 size 32x32
      Appearance <- "Barcode506"
   Circle "Circle_8" at 102,279 size 32x32
      Appearance <- "Barcode515"
   Circle "Circle_11" at 166,164 size 32x32
      Appearance <- "Barcode498"
   Circle "Circle_12" at 166,224 size 32x32
      Appearance <- "Barcode507"
   Circle "Circle_13" at 166,279 size 32x32
      Appearance <- "Barcode516"
   Circle "Circle_16" at 227,165 size 32x32
      Appearance <- "Barcode499"
   Circle "Circle_17" at 230,224 size 32x32
      Appearance <- "Barcode508"
   Circle "Circle_18" at 230,279 size 32x32
      Appearance <- "Barcode517"
   Circle "Circle_21" at 294,164 size 32x32
      Appearance <- "Barcode500"
   Circle "Circle_22" at 294,224 size 32x32
      Appearance <- "Barcode509"
   Circle "Circle_23" at 294,279 size 32x32
      Appearance <- "Barcode518"
   Circle "Circle_26" at 358,164 size 32x32
      Appearance <- "Barcode501"
   Circle "Circle_27" at 358,225 size 32x32
      Appearance <- "Barcode510"
   Circle "Circle_28" at 358,279 size 32x32
      Appearance <- "Barcode519"
   Circle "Circle_31" at 422,164 size 32x32
      Appearance <- "Barcode502"
   Circle "Circle_32" at 422,224 size 32x32
      Appearance <- "Barcode511"
   Circle "Circle_33" at 422,279 size 32x32
      Appearance <- "Barcode520"
   Circle "Circle_36" at 486,164 size 32x32
      Appearance <- "Barcode503"
   Circle "Circle_37" at 486,224 size 32x32
      Appearance <- "Barcode512"
   Circle "Circle_41" at 550,163 size 32x32
      Appearance <- "Barcode504"
   Circle "Circle_42" at 550,224 size 32x32
      Appearance <- "Barcode513"
   GraphicView "Template_Graphic view_3" at 8,6 size 70x68; Picture "KMUTNB-Photoroom"
   GraphicView "Template_Graphic view_5" at 657,59 size 104x124; Picture "channels4_profile-Photoroom"
   Button "Button_5" at 633,292 size 64x24; TextOff 'Back'
      on Click: ActivateScreen("Screen_11", 0)
   GraphicView "Template_Graphic view_4" at 736,255 size 28x26; Picture "NEW_HOME"
   GraphicView "Template_Graphic view_2" at 650,253 size 28x27; Picture "play"
   GraphicView "Template_Graphic view_6" at 638,296 size 20x17; Picture "previous-track"
   Button "Button_1" at 623,245 size 80x42; TextOff 'Text'
      on Press: SetTag("มีการปุ่มกดยืนยัน", 1)
      on Release: SetTag("มีการปุ่มกดยืนยัน", 0)
      on Activate: "Storage"()
   Button "Button_3" at 707,246 size 80x42; TextOn 'LOGOUT'; TextOff 'Text'
      on Activate: function_f23ef4c9(); ActivateScreen("1_OVERVIEW_1", 0)
   TextField "Text field_49" at 734,229 size 32x14; Text 'HOME'
   TextField "Text field_50" at 625,229 size 95x16; Text 'Simmulation Conveyor'

VB script "Retrieval"
   'Tip:
   ' 1. Use the <CTRL+SPACE> or <CTRL+I> shortcut to open a list of all objects and functions
   ' 2. Write the code using the HMI Runtime object.
   '  Example: HmiRuntime.Screens("Screen_1").
   ' 3. Use the <CTRL+J> shortcut to create an object reference.
   'Write the code as of this position:
   Dim u, p, nm
   u = SmartTags("Selected_URL")
   p = InStrRev(u, "/")
   nm = Replace(Mid(u, p + 1), ".html", "")
   SmartTags("Video_URL") = Left(u, p) & "player.html#c=" & nm & "&t=" & (Hour(Now)*3600 + Minute(Now)*60 + Second(Now))

VB script "Storage"
   'Tip:
   ' 1. Use the <CTRL+SPACE> or <CTRL+I> shortcut to open a list of all objects and functions
   ' 2. Write the code using the HMI Runtime object.
   '  Example: HmiRuntime.Screens("Screen_1").
   ' 3. Use the <CTRL+J> shortcut to create an object reference.
   'Write the code as of this position:
   Dim code
   code = UCase(Trim(SmartTags("Expected/Value_All_V")))
   If code = "" Then Exit Sub
   SmartTags("Video_URL") = "file:///C:/ASRS_Video/Storage/player.html#c=" & code & "&t=" & (Hour(Now)*3600 + Minute(Now)*60 + Second(Now))
   bec8f1e5-2ab1-45f6-ad91-1d37c469eb91 Screen_1, 0

VB script "Conveyor"
   'Tip:
   ' 1. Use the <CTRL+SPACE> or <CTRL+I> shortcut to open a list of all objects and functions
   ' 2. Write the code using the HMI Runtime object.
   '  Example: HmiRuntime.Screens("Screen_1").
   ' 3. Use the <CTRL+J> shortcut to create an object reference.
   'Write the code as of this position:
   SmartTags("Video_URL") = "file:///C:/ASRS_Video/Storage/player.html#c=conveyor&t=" & (Hour(Now)*3600 + Minute(Now)*60 + Second(Now))

VB script "Test2"
   'Tip:
   ' 1. Use the <CTRL+SPACE> or <CTRL+I> shortcut to open a list of all objects and functions
   ' 2. Write the code using the HMI Runtime object.
   '  Example: HmiRuntime.Screens("Screen_1").
   ' 3. Use the <CTRL+J> shortcut to create an object reference.
   'Write the code as of this position:
   Dim Barcode
   Dim shell
   
   Barcode = SmartTags("Expected/Value_All_V")
   
   Set shell = CreateObject("WScript.Shell")
   
   If Barcode = "A001" Then
       shell.Run "C:\Users\poh25\Videos\VMed 520box\Full-All-001.mp4"
   
   ElseIf Barcode = "A002" Then
       shell.Run "C:\Users\poh25\Videos\mini\A002.mp4"
   
   ElseIf Barcode = "A003" Then
       shell.Run "C:\Users\poh25\Videos\mini\A003.mp4"
   
   ElseIf Barcode = "A004" Then
       shell.Run "C:\Users\poh25\Videos\mini\A004.mp4"
   
   ElseIf Barcode = "A005" Then
       shell.Run "C:\Users\poh25\Videos\mini\A005.mp4"
   
   ElseIf Barcode = "A006" Then
       shell.Run "C:\Users\poh25\Videos\mini\A006.mp4"
   
   ElseIf Barcode = "A007" Then
       shell.Run "C:\Users\poh25\Videos\mini\A007.mp4"
   
   ElseIf Barcode = "A008" Then
       shell.Run "C:\Users\poh25\Videos\mini\A008.mp4"
   
   ElseIf Barcode = "A009" Then
       shell.Run "C:\Users\poh25\Videos\mini\A009.mp4"
   
   ElseIf Barcode = "A010" Then
       shell.Run "C:\Users\poh25\Videos\mini\A010.mp4"
   
   ElseIf Barcode = "A011" Then
       shell.Run "C:\Users\poh25\Videos\mini\A011.mp4"
   
   ElseIf Barcode = "A012" Then
       shell.Run "C:\Users\poh25\Videos\mini\A012.mp4"
   
   ElseIf Barcode = "A013" Then
       shell.Run "C:\Users\poh25\Videos\mini\A013.mp4"
   
   ElseIf Barcode = "A014" Then
       shell.Run "C:\Users\poh25\Videos\mini\A014.mp4"
   
   ElseIf Barcode = "A015" Then
       shell.Run "C:\Users\poh25\Videos\mini\A015.mp4"
   
   ElseIf Barcode = "A016" Then
       shell.Run "C:\Users\poh25\Videos\mini\A016.mp4"
   
   ElseIf Barcode = "A017" Then
       shell.Run "C:\Users\poh25\Videos\mini\A017.mp4"
   
   ElseIf Barcode = "A018" Then
       shell.Run "C:\Users\poh25\Videos\mini\A018.mp4"
   
   ElseIf Barcode = "A019" Then
       shell.Run "C:\Users\poh25\Videos\mini\A019.mp4"
   
   ElseIf Barcode = "A020" Then
       shell.Run "C:\Users\poh25\Videos\mini\A020.mp4"
   
   ElseIf Barcode = "A021" Then
       shell.Run "C:\Users\poh25\Videos\mini\A021.mp4"
   
   ElseIf Barcode = "A022" Then
       shell.Run "C:\Users\poh25\Videos\mini\A022.mp4"
   
   ElseIf Barcode = "A023" Then
       shell.Run "C:\Users\poh25\Videos\mini\A023.mp4"
   
   ElseIf Barcode = "A024" Then
       shell.Run "C:\Users\poh25\Videos\mini\A024.mp4"
   
   ElseIf Barcode = "A025" Then
       shell.Run "C:\Users\poh25\Videos\mini\A025.mp4"
   
   ElseIf Barcode = "A026" Then
       shell.Run "C:\Users\poh25\Videos\mini\A026.mp4"
   
   ElseIf Barcode = "A027" Then
       shell.Run "C:\Users\poh25\Videos\mini\A027.mp4"
   
   ElseIf Barcode = "A028" Then
       shell.Run "C:\Users\poh25\Videos\mini\A028.mp4"
   
   ElseIf Barcode = "A029" Then
       shell.Run "C:\Users\poh25\Videos\mini\A029.mp4"
   
   ElseIf Barcode = "A030" Then
       shell.Run "C:\Users\poh25\Videos\mini\A030.mp4"
   
   ElseIf Barcode = "A031" Then
       shell.Run "C:\Users\poh25\Videos\mini\A031.mp4"
   
   ElseIf Barcode = "A032" Then
       shell.Run "C:\Users\poh25\Videos\mini\A032.mp4"
   
   ElseIf Barcode = "A033" Then
       shell.Run "C:\Users\poh25\Videos\mini\A033.mp4"
   
   ElseIf Barcode = "A034" Then
       shell.Run "C:\Users\poh25\Videos\mini\A034.mp4"
   
   ElseIf Barcode = "A035" Then
       shell.Run "C:\Users\poh25\Videos\mini\A035.mp4"
   
   ElseIf Barcode = "A036" Then
       shell.Run "C:\Users\poh25\Videos\mini\A036.mp4"
   
   ElseIf Barcode = "A037" Then
       shell.Run "C:\Users\poh25\Videos\mini\A037.mp4"
   
   ElseIf Barcode = "A038" Then
       shell.Run "C:\Users\poh25\Videos\mini\A038.mp4"
   
   ElseIf Barcode = "A039" Then
       shell.Run "C:\Users\poh25\Videos\mini\A039.mp4"
   
   ElseIf Barcode = "A040" Then
       shell.Run "C:\Users\poh25\Videos\mini\A040.mp4"
   
   ElseIf Barcode = "A041" Then
       shell.Run "C:\Users\poh25\Videos\mini\A041.mp4"
   
   ElseIf Barcode = "A042" Then
       shell.Run "C:\Users\poh25\Videos\mini\A042.mp4"
   
   ElseIf Barcode = "A043" Then
       shell.Run "C:\Users\poh25\Videos\mini\A043.mp4"
   
   ElseIf Barcode = "A044" Then
       shell.Run "C:\Users\poh25\Videos\mini\A044.mp4"
   
   ElseIf Barcode = "A045" Then
       shell.Run "C:\Users\poh25\Videos\mini\A045.mp4"
   
   ElseIf Barcode = "A046" Then
       shell.Run "C:\Users\poh25\Videos\mini\A046.mp4"
   
   ElseIf Barcode = "A047" Then
       shell.Run "C:\Users\poh25\Videos\mini\A047.mp4"
   
   ElseIf Barcode = "A048" Then
       shell.Run "C:\Users\poh25\Videos\mini\A048.mp4"
   
   ElseIf Barcode = "A049" Then
       shell.Run "C:\Users\poh25\Videos\mini\A049.mp4"
   
   ElseIf Barcode = "A050" Then
       shell.Run "C:\Users\poh25\Videos\mini\A050.mp4"
   
   ElseIf Barcode = "A051" Then
       shell.Run "C:\Users\poh25\Videos\mini\A051.mp4"
   
   ElseIf Barcode = "A052" Then
       shell.Run "C:\Users\poh25\Videos\mini\A052.mp4"
   
   ElseIf Barcode = "A053" Then
       shell.Run "C:\Users\poh25\Videos\mini\A053.mp4"
   
   ElseIf Barcode = "A054" Then
       shell.Run "C:\Users\poh25\Videos\mini\A054.mp4"
   
   ElseIf Barcode = "A055" Then
       shell.Run "C:\Users\poh25\Videos\mini\A055.mp4"
   
   ElseIf Barcode = "A056" Then
       shell.Run "C:\Users\poh25\Videos\mini\A056.mp4"
   
   ElseIf Barcode = "A057" Then
       shell.Run "C:\Users\poh25\Videos\mini\A057.mp4"
   
   ElseIf Barcode = "A058" Then
       shell.Run "C:\Users\poh25\Videos\mini\A058.mp4"
   
   ElseIf Barcode = "A059" Then
       shell.Run "C:\Users\poh25\Videos\mini\A059.mp4"
   
   ElseIf Barcode = "A060" Then
       shell.Run "C:\Users\poh25\Videos\mini\A060.mp4"
   
   ElseIf Barcode = "A061" Then
       shell.Run "C:\Users\poh25\Videos\mini\A061.mp4"
   
   ElseIf Barcode = "A062" Then
       shell.Run "C:\Users\poh25\Videos\mini\A062.mp4"
   
   ElseIf Barcode = "A063" Then
       shell.Run "C:\Users\poh25\Videos\mini\A063.mp4"
   
   ElseIf Barcode = "A064" Then
       shell.Run "C:\Users\poh25\Videos\mini\A064.mp4"
   
   ElseIf Barcode = "A065" Then
       shell.Run "C:\Users\poh25\Videos\mini\A065.mp4"
   
   ElseIf Barcode = "A066" Then
       shell.Run "C:\Users\poh25\Videos\mini\A066.mp4"
   
   ElseIf Barcode = "A067" Then
       shell.Run "C:\Users\poh25\Videos\mini\A067.mp4"
   
   ElseIf Barcode = "A068" Then
       shell.Run "C:\Users\poh25\Videos\mini\A068.mp4"
   
   ElseIf Barcode = "A069" Then
       shell.Run "C:\Users\poh25\Videos\mini\A069.mp4"
   
   ElseIf Barcode = "A070" Then
       shell.Run "C:\Users\poh25\Videos\mini\A070.mp4"
   
   ElseIf Barcode = "A071" Then
       shell.Run "C:\Users\poh25\Videos\mini\A071.mp4"
   
   ElseIf Barcode = "A072" Then
       shell.Run "C:\Users\poh25\Videos\mini\A072.mp4"
   
   ElseIf Barcode = "A073" Then
       shell.Run "C:\Users\poh25\Videos\mini\A073.mp4"
   
   ElseIf Barcode = "A074" Then
       shell.Run "C:\Users\poh25\Videos\mini\A074.mp4"
   
   ElseIf Barcode = "A075" Then
       shell.Run "C:\Users\poh25\Videos\mini\A075.mp4"
   
   ElseIf Barcode = "A076" Then
       shell.Run "C:\Users\poh25\Videos\mini\A076.mp4"
   
   ElseIf Barcode = "A077" Then
       shell.Run "C:\Users\poh25\Videos\mini\A077.mp4"
   
   ElseIf Barcode = "A078" Then
       shell.Run "C:\Users\poh25\Videos\mini\A078.mp4"
   
   ElseIf Barcode = "A079" Then
       shell.Run "C:\Users\poh25\Videos\mini\A079.mp4"
   
   ElseIf Barcode = "A080" Then
       shell.Run "C:\Users\poh25\Videos\mini\A080.mp4"
   
   ElseIf Barcode = "A081" Then
       shell.Run "C:\Users\poh25\Videos\mini\A081.mp4"
   
   ElseIf Barcode = "A082" Then
       shell.Run "C:\Users\poh25\Videos\mini\A082.mp4"
   
   ElseIf Barcode = "A083" Then
       shell.Run "C:\Users\poh25\Videos\mini\A083.mp4"
   
   ElseIf Barcode = "A084" Then
       shell.Run "C:\Users\poh25\Videos\mini\A084.mp4"
   
   ElseIf Barcode = "A085" Then
       shell.Run "C:\Users\poh25\Videos\mini\A085.mp4"
   
   ElseIf Barcode = "A086" Then
       shell.Run "C:\Users\poh25\Videos\mini\A086.mp4"
   
   ElseIf Barcode = "A087" Then
       shell.Run "C:\Users\poh25\Videos\mini\A087.mp4"
   
   ElseIf Barcode = "A088" Then
       shell.Run "C:\Users\poh25\Videos\mini\A088.mp4"
   
   ElseIf Barcode = "A089" Then
       shell.Run "C:\Users\poh25\Videos\mini\A089.mp4"
   
   ElseIf Barcode = "A090" Then
       shell.Run "C:\Users\poh25\Videos\mini\A090.mp4"
   
   ElseIf Barcode = "A091" Then
       shell.Run "C:\Users\poh25\Videos\mini\A091.mp4"
   
   ElseIf Barcode = "A092" Then
       shell.Run "C:\Users\poh25\Videos\mini\A092.mp4"
   
   ElseIf Barcode = "A093" Then
       shell.Run "C:\Users\poh25\Videos\mini\A093.mp4"
   
   ElseIf Barcode = "A094" Then
       shell.Run "C:\Users\poh25\Videos\mini\A094.mp4"
   
   ElseIf Barcode = "A095" Then
       shell.Run "C:\Users\poh25\Videos\mini\A095.mp4"
   
   ElseIf Barcode = "A096" Then
       shell.Run "C:\Users\poh25\Videos\mini\A096.mp4"
   
   ElseIf Barcode = "A097" Then
       shell.Run "C:\Users\poh25\Videos\mini\A097.mp4"
   
   ElseIf Barcode = "A098" Then
       shell.Run "C:\Users\poh25\Videos\mini\A098.mp4"
   
   ElseIf Barcode = "A099" Then
       shell.Run "C:\Users\poh25\Videos\mini\A099.mp4"
   
   ElseIf Barcode = "A100" Then
       shell.Run "C:\Users\poh25\Videos\mini\A100.mp4"
   
   ElseIf Barcode = "B001" Then
       shell.Run "C:\Users\poh25\Videos\mini\B001.mp4"
   
   ElseIf Barcode = "B002" Then
       shell.Run "C:\Users\poh25\Videos\mini\B002.mp4"
   
   ElseIf Barcode = "B003" Then
       shell.Run "C:\Users\poh25\Videos\mini\B003.mp4"
   
   ElseIf Barcode = "B004" Then
       shell.Run "C:\Users\poh25\Videos\mini\B004.mp4"
   
   ElseIf Barcode = "B005" Then
       shell.Run "C:\Users\poh25\Videos\mini\B005.mp4"
   
   ElseIf Barcode = "B006" Then
       shell.Run "C:\Users\poh25\Videos\mini\B006.mp4"
   
   ElseIf Barcode = "B007" Then
       shell.Run "C:\Users\poh25\Videos\mini\B007.mp4"
   
   ElseIf Barcode = "B008" Then
       shell.Run "C:\Users\poh25\Videos\mini\B008.mp4"
   
   ElseIf Barcode = "B009" Then
       shell.Run "C:\Users\poh25\Videos\mini\B009.mp4"
   
   ElseIf Barcode = "B010" Then
       shell.Run "C:\Users\poh25\Videos\mini\B010.mp4"
   
   ElseIf Barcode = "B011" Then
       shell.Run "C:\Users\poh25\Videos\mini\B011.mp4"
   
   ElseIf Barcode = "B012" Then
       shell.Run "C:\Users\poh25\Videos\mini\B012.mp4"
   
   ElseIf Barcode = "B013" Then
       shell.Run "C:\Users\poh25\Videos\mini\B013.mp4"
   
   ElseIf Barcode = "B014" Then
       shell.Run "C:\Users\poh25\Videos\mini\B014.mp4"
   
   ElseIf Barcode = "B015" Then
       shell.Run "C:\Users\poh25\Videos\mini\B015.mp4"
   
   ElseIf Barcode = "B016" Then
       shell.Run "C:\Users\poh25\Videos\mini\B016.mp4"
   
   ElseIf Barcode = "B017" Then
       shell.Run "C:\Users\poh25\Videos\mini\B017.mp4"
   
   ElseIf Barcode = "B018" Then
       shell.Run "C:\Users\poh25\Videos\mini\B018.mp4"
   
   ElseIf Barcode = "B019" Then
       shell.Run "C:\Users\poh25\Videos\mini\B019.mp4"
   
   ElseIf Barcode = "B020" Then
       shell.Run "C:\Users\poh25\Videos\mini\B020.mp4"
   
   ElseIf Barcode = "B021" Then
       shell.Run "C:\Users\poh25\Videos\mini\B021.mp4"
   
   ElseIf Barcode = "B022" Then
       shell.Run "C:\Users\poh25\Videos\mini\B022.mp4"
   
   ElseIf Barcode = "B023" Then
       shell.Run "C:\Users\poh25\Videos\mini\B023.mp4"
   
   ElseIf Barcode = "B024" Then
       shell.Run "C:\Users\poh25\Videos\mini\B024.mp4"
   
   ElseIf Barcode = "B025" Then
       shell.Run "C:\Users\poh25\Videos\mini\B025.mp4"
   
   ElseIf Barcode = "B026" Then
       shell.Run "C:\Users\poh25\Videos\mini\B026.mp4"
   
   ElseIf Barcode = "B027" Then
       shell.Run "C:\Users\poh25\Videos\mini\B027.mp4"
   
   ElseIf Barcode = "B028" Then
       shell.Run "C:\Users\poh25\Videos\mini\B028.mp4"
   
   ElseIf Barcode = "B029" Then
       shell.Run "C:\Users\poh25\Videos\mini\B029.mp4"
   
   ElseIf Barcode = "B030" Then
       shell.Run "C:\Users\poh25\Videos\mini\B030.mp4"
   
   ElseIf Barcode = "B031" Then
       shell.Run "C:\Users\poh25\Videos\mini\B031.mp4"
   
   ElseIf Barcode = "B032" Then
       shell.Run "C:\Users\poh25\Videos\mini\B032.mp4"
   
   ElseIf Barcode = "B033" Then
       shell.Run "C:\Users\poh25\Videos\mini\B033.mp4"
   
   ElseIf Barcode = "B034" Then
       shell.Run "C:\Users\poh25\Videos\mini\B034.mp4"
   
   ElseIf Barcode = "B035" Then
       shell.Run "C:\Users\poh25\Videos\mini\B035.mp4"
   
   ElseIf Barcode = "B036" Then
       shell.Run "C:\Users\poh25\Videos\mini\B036.mp4"
   
   ElseIf Barcode = "B037" Then
       shell.Run "C:\Users\poh25\Videos\mini\B037.mp4"
   
   ElseIf Barcode = "B038" Then
       shell.Run "C:\Users\poh25\Videos\mini\B038.mp4"
   
   ElseIf Barcode = "B039" Then
       shell.Run "C:\Users\poh25\Videos\mini\B039.mp4"
   
   ElseIf Barcode = "B040" Then
       shell.Run "C:\Users\poh25\Videos\mini\B040.mp4"
   
   ElseIf Barcode = "B041" Then
       shell.Run "C:\Users\poh25\Videos\mini\B041.mp4"
   
   ElseIf Barcode = "B042" Then
       shell.Run "C:\Users\poh25\Videos\mini\B042.mp4"
   
   ElseIf Barcode = "B043" Then
       shell.Run "C:\Users\poh25\Videos\mini\B043.mp4"
   
   ElseIf Barcode = "B044" Then
       shell.Run "C:\Users\poh25\Videos\mini\B044.mp4"
   
   ElseIf Barcode = "B045" Then
       shell.Run "C:\Users\poh25\Videos\mini\B045.mp4"
   
   ElseIf Barcode = "B046" Then
       shell.Run "C:\Users\poh25\Videos\mini\B046.mp4"
   
   ElseIf Barcode = "B047" Then
       shell.Run "C:\Users\poh25\Videos\mini\B047.mp4"
   
   ElseIf Barcode = "B048" Then
       shell.Run "C:\Users\poh25\Videos\mini\B048.mp4"
   
   ElseIf Barcode = "B049" Then
       shell.Run "C:\Users\poh25\Videos\mini\B049.mp4"
   
   ElseIf Barcode = "B050" Then
       shell.Run "C:\Users\poh25\Videos\mini\B050.mp4"
   
   ElseIf Barcode = "B051" Then
       shell.Run "C:\Users\poh25\Videos\mini\B051.mp4"
   
   ElseIf Barcode = "B052" Then
       shell.Run "C:\Users\poh25\Videos\mini\B052.mp4"
   
   ElseIf Barcode = "B053" Then
       shell.Run "C:\Users\poh25\Videos\mini\B053.mp4"
   
   ElseIf Barcode = "B054" Then
       shell.Run "C:\Users\poh25\Videos\mini\B054.mp4"
   
   ElseIf Barcode = "B055" Then
       shell.Run "C:\Users\poh25\Videos\mini\B055.mp4"
   
   ElseIf Barcode = "B056" Then
       shell.Run "C:\Users\poh25\Videos\mini\B056.mp4"
   
   ElseIf Barcode = "B057" Then
       shell.Run "C:\Users\poh25\Videos\mini\B057.mp4"
   
   ElseIf Barcode = "B058" Then
       shell.Run "C:\Users\poh25\Videos\mini\B058.mp4"
   
   ElseIf Barcode = "B059" Then
       shell.Run "C:\Users\poh25\Videos\mini\B059.mp4"
   
   ElseIf Barcode = "B060" Then
       shell.Run "C:\Users\poh25\Videos\mini\B060.mp4"
   
   ElseIf Barcode = "B061" Then
       shell.Run "C:\Users\poh25\Videos\mini\B061.mp4"
   
   ElseIf Barcode = "B062" Then
       shell.Run "C:\Users\poh25\Videos\mini\B062.mp4"
   
   ElseIf Barcode = "B063" Then
       shell.Run "C:\Users\poh25\Videos\mini\B063.mp4"
   
   ElseIf Barcode = "B064" Then
       shell.Run "C:\Users\poh25\Videos\mini\B064.mp4"
   
   ElseIf Barcode = "B065" Then
       shell.Run "C:\Users\poh25\Videos\mini\B065.mp4"
   
   ElseIf Barcode = "B066" Then
       shell.Run "C:\Users\poh25\Videos\mini\B066.mp4"
   
   ElseIf Barcode = "B067" Then
       shell.Run "C:\Users\poh25\Videos\mini\B067.mp4"
   
   ElseIf Barcode = "B068" Then
       shell.Run "C:\Users\poh25\Videos\mini\B068.mp4"
   
   ElseIf Barcode = "B069" Then
       shell.Run "C:\Users\poh25\Videos\mini\B069.mp4"
   
   ElseIf Barcode = "B070" Then
       shell.Run "C:\Users\poh25\Videos\mini\B070.mp4"
   
   ElseIf Barcode = "B071" Then
       shell.Run "C:\Users\poh25\Videos\mini\B071.mp4"
   
   ElseIf Barcode = "B072" Then
       shell.Run "C:\Users\poh25\Videos\mini\B072.mp4"
   
   ElseIf Barcode = "B073" Then
       shell.Run "C:\Users\poh25\Videos\mini\B073.mp4"
   
   ElseIf Barcode = "B074" Then
       shell.Run "C:\Users\poh25\Videos\mini\B074.mp4"
   
   ElseIf Barcode = "B075" Then
       shell.Run "C:\Users\poh25\Videos\mini\B075.mp4"
   
   ElseIf Barcode = "B076" Then
       shell.Run "C:\Users\poh25\Videos\mini\B076.mp4"
   
   ElseIf Barcode = "B077" Then
       shell.Run "C:\Users\poh25\Videos\mini\B077.mp4"
   
   ElseIf Barcode = "B078" Then
       shell.Run "C:\Users\poh25\Videos\mini\B078.mp4"
   
   ElseIf Barcode = "B079" Then
       shell.Run "C:\Users\poh25\Videos\mini\B079.mp4"
   
   ElseIf Barcode = "B080" Then
       shell.Run "C:\Users\poh25\Videos\mini\B080.mp4"
   
   ElseIf Barcode = "B081" Then
       shell.Run "C:\Users\poh25\Videos\mini\B081.mp4"
   
   ElseIf Barcode = "B082" Then
       shell.Run "C:\Users\poh25\Videos\mini\B082.mp4"
   
   ElseIf Barcode = "B083" Then
       shell.Run "C:\Users\poh25\Videos\mini\B083.mp4"
   
   ElseIf Barcode = "B084" Then
       shell.Run "C:\Users\poh25\Videos\mini\B084.mp4"
   
   ElseIf Barcode = "B085" Then
       shell.Run "C:\Users\poh25\Videos\mini\B085.mp4"
   
   ElseIf Barcode = "B086" Then
       shell.Run "C:\Users\poh25\Videos\mini\B086.mp4"
   
   ElseIf Barcode = "B087" Then
       shell.Run "C:\Users\poh25\Videos\mini\B087.mp4"
   
   ElseIf Barcode = "B088" Then
       shell.Run "C:\Users\poh25\Videos\mini\B088.mp4"
   
   ElseIf Barcode = "B089" Then
       shell.Run "C:\Users\poh25\Videos\mini\B089.mp4"
   
   ElseIf Barcode = "B090" Then
       shell.Run "C:\Users\poh25\Videos\mini\B090.mp4"
   
   ElseIf Barcode = "B091" Then
       shell.Run "C:\Users\poh25\Videos\mini\B091.mp4"
   
   ElseIf Barcode = "B092" Then
       shell.Run "C:\Users\poh25\Videos\mini\B092.mp4"
   
   ElseIf Barcode = "B093" Then
       shell.Run "C:\Users\poh25\Videos\mini\B093.mp4"
   
   ElseIf Barcode = "B094" Then
       shell.Run "C:\Users\poh25\Videos\mini\B094.mp4"
   
   ElseIf Barcode = "B095" Then
       shell.Run "C:\Users\poh25\Videos\mini\B095.mp4"
   
   ElseIf Barcode = "B096" Then
       shell.Run "C:\Users\poh25\Videos\mini\B096.mp4"
   
   ElseIf Barcode = "B097" Then
       shell.Run "C:\Users\poh25\Videos\mini\B097.mp4"
   
   ElseIf Barcode = "B098" Then
       shell.Run "C:\Users\poh25\Videos\mini\B098.mp4"
   
   ElseIf Barcode = "B099" Then
       shell.Run "C:\Users\poh25\Videos\mini\B099.mp4"
   
   ElseIf Barcode = "B100" Then
       shell.Run "C:\Users\poh25\Videos\mini\B100.mp4"
   
   ElseIf Barcode = "C001" Then
       shell.Run "C:\Users\poh25\Videos\mini\C001.mp4"
   
   ElseIf Barcode = "C002" Then
       shell.Run "C:\Users\poh25\Videos\mini\C002.mp4"
   
   ElseIf Barcode = "C003" Then
       shell.Run "C:\Users\poh25\Videos\mini\C003.mp4"
   
   ElseIf Barcode = "C004" Then
       shell.Run "C:\Users\poh25\Videos\mini\C004.mp4"
   
   ElseIf Barcode = "C005" Then
       shell.Run "C:\Users\poh25\Videos\mini\C005.mp4"
   
   ElseIf Barcode = "C006" Then
       shell.Run "C:\Users\poh25\Videos\mini\C006.mp4"
   
   ElseIf Barcode = "C007" Then
       shell.Run "C:\Users\poh25\Videos\mini\C007.mp4"
   
   ElseIf Barcode = "C008" Then
       shell.Run "C:\Users\poh25\Videos\mini\C008.mp4"
   
   ElseIf Barcode = "C009" Then
       shell.Run "C:\Users\poh25\Videos\mini\C009.mp4"
   
   ElseIf Barcode = "C010" Then
       shell.Run "C:\Users\poh25\Videos\mini\C010.mp4"
   
   ElseIf Barcode = "C011" Then
       shell.Run "C:\Users\poh25\Videos\mini\C011.mp4"
   
   ElseIf Barcode = "C012" Then
       shell.Run "C:\Users\poh25\Videos\mini\C012.mp4"
   
   ElseIf Barcode = "C013" Then
       shell.Run "C:\Users\poh25\Videos\mini\C013.mp4"
   
   ElseIf Barcode = "C014" Then
       shell.Run "C:\Users\poh25\Videos\mini\C014.mp4"
   
   ElseIf Barcode = "C015" Then
       shell.Run "C:\Users\poh25\Videos\mini\C015.mp4"
   
   ElseIf Barcode = "C016" Then
       shell.Run "C:\Users\poh25\Videos\mini\C016.mp4"
   
   ElseIf Barcode = "C017" Then
       shell.Run "C:\Users\poh25\Videos\mini\C017.mp4"
   
   ElseIf Barcode = "C018" Then
       shell.Run "C:\Users\poh25\Videos\mini\C018.mp4"
   
   ElseIf Barcode = "C019" Then
       shell.Run "C:\Users\poh25\Videos\mini\C019.mp4"
   
   ElseIf Barcode = "C020" Then
       shell.Run "C:\Users\poh25\Videos\mini\C020.mp4"
   
   ElseIf Barcode = "C021" Then
       shell.Run "C:\Users\poh25\Videos\mini\C021.mp4"
   
   ElseIf Barcode = "C022" Then
       shell.Run "C:\Users\poh25\Videos\mini\C022.mp4"
   
   ElseIf Barcode = "C023" Then
       shell.Run "C:\Users\poh25\Videos\mini\C023.mp4"
   
   ElseIf Barcode = "C024" Then
       shell.Run "C:\Users\poh25\Videos\mini\C024.mp4"
   
   ElseIf Barcode = "C025" Then
       shell.Run "C:\Users\poh25\Videos\mini\C025.mp4"
   
   ElseIf Barcode = "C026" Then
       shell.Run "C:\Users\poh25\Videos\mini\C026.mp4"
   
   ElseIf Barcode = "C027" Then
       shell.Run "C:\Users\poh25\Videos\mini\C027.mp4"
   
   ElseIf Barcode = "C028" Then
       shell.Run "C:\Users\poh25\Videos\mini\C028.mp4"
   
   ElseIf Barcode = "C029" Then
       shell.Run "C:\Users\poh25\Videos\mini\C029.mp4"
   
   ElseIf Barcode = "C030" Then
       shell.Run "C:\Users\poh25\Videos\mini\C030.mp4"
   
   ElseIf Barcode = "C031" Then
       shell.Run "C:\Users\poh25\Videos\mini\C031.mp4"
   
   ElseIf Barcode = "C032" Then
       shell.Run "C:\Users\poh25\Videos\mini\C032.mp4"
   
   ElseIf Barcode = "C033" Then
       shell.Run "C:\Users\poh25\Videos\mini\C033.mp4"
   
   ElseIf Barcode = "C034" Then
       shell.Run "C:\Users\poh25\Videos\mini\C034.mp4"
   
   ElseIf Barcode = "C035" Then
       shell.Run "C:\Users\poh25\Videos\mini\C035.mp4"
   
   ElseIf Barcode = "C036" Then
       shell.Run "C:\Users\poh25\Videos\mini\C036.mp4"
   
   ElseIf Barcode = "C037" Then
       shell.Run "C:\Users\poh25\Videos\mini\C037.mp4"
   
   ElseIf Barcode = "C038" Then
       shell.Run "C:\Users\poh25\Videos\mini\C038.mp4"
   
   ElseIf Barcode = "C039" Then
       shell.Run "C:\Users\poh25\Videos\mini\C039.mp4"
   
   ElseIf Barcode = "C040" Then
       shell.Run "C:\Users\poh25\Videos\mini\C040.mp4"
   
   ElseIf Barcode = "C041" Then
       shell.Run "C:\Users\poh25\Videos\mini\C041.mp4"
   
   ElseIf Barcode = "C042" Then
       shell.Run "C:\Users\poh25\Videos\mini\C042.mp4"
   
   ElseIf Barcode = "C043" Then
       shell.Run "C:\Users\poh25\Videos\mini\C043.mp4"
   
   ElseIf Barcode = "C044" Then
       shell.Run "C:\Users\poh25\Videos\mini\C044.mp4"
   
   ElseIf Barcode = "C045" Then
       shell.Run "C:\Users\poh25\Videos\mini\C045.mp4"
   
   ElseIf Barcode = "C046" Then
       shell.Run "C:\Users\poh25\Videos\mini\C046.mp4"
   
   ElseIf Barcode = "C047" Then
       shell.Run "C:\Users\poh25\Videos\mini\C047.mp4"
   
   ElseIf Barcode = "C048" Then
       shell.Run "C:\Users\poh25\Videos\mini\C048.mp4"
   
   ElseIf Barcode = "C049" Then
       shell.Run "C:\Users\poh25\Videos\mini\C049.mp4"
   
   ElseIf Barcode = "C050" Then
       shell.Run "C:\Users\poh25\Videos\mini\C050.mp4"
   
   ElseIf Barcode = "C051" Then
       shell.Run "C:\Users\poh25\Videos\mini\C051.mp4"
   
   ElseIf Barcode = "C052" Then
       shell.Run "C:\Users\poh25\Videos\mini\C052.mp4"
   
   ElseIf Barcode = "C053" Then
       shell.Run "C:\Users\poh25\Videos\mini\C053.mp4"
   
   ElseIf Barcode = "C054" Then
       shell.Run "C:\Users\poh25\Videos\mini\C054.mp4"
   
   ElseIf Barcode = "C055" Then
       shell.Run "C:\Users\poh25\Videos\mini\C055.mp4"
   
   ElseIf Barcode = "C056" Then
       shell.Run "C:\Users\poh25\Videos\mini\C056.mp4"
   
   ElseIf Barcode = "C057" Then
       shell.Run "C:\Users\poh25\Videos\mini\C057.mp4"
   
   ElseIf Barcode = "C058" Then
       shell.Run "C:\Users\poh25\Videos\mini\C058.mp4"
   
   ElseIf Barcode = "C059" Then
       shell.Run "C:\Users\poh25\Videos\mini\C059.mp4"
   
   ElseIf Barcode = "C060" Then
       shell.Run "C:\Users\poh25\Videos\mini\C060.mp4"
   
   ElseIf Barcode = "C061" Then
       shell.Run "C:\Users\poh25\Videos\mini\C061.mp4"
   
   ElseIf Barcode = "C062" Then
       shell.Run "C:\Users\poh25\Videos\mini\C062.mp4"
   
   ElseIf Barcode = "C063" Then
       shell.Run "C:\Users\poh25\Videos\mini\C063.mp4"
   
   ElseIf Barcode = "C064" Then
       shell.Run "C:\Users\poh25\Videos\mini\C064.mp4"
   
   ElseIf Barcode = "C065" Then
       shell.Run "C:\Users\poh25\Videos\mini\C065.mp4"
   
   ElseIf Barcode = "C066" Then
       shell.Run "C:\Users\poh25\Videos\mini\C066.mp4"
   
   ElseIf Barcode = "C067" Then
       shell.Run "C:\Users\poh25\Videos\mini\C067.mp4"
   
   ElseIf Barcode = "C068" Then
       shell.Run "C:\Users\poh25\Videos\mini\C068.mp4"
   
   ElseIf Barcode = "C069" Then
       shell.Run "C:\Users\poh25\Videos\mini\C069.mp4"
   
   ElseIf Barcode = "C070" Then
       shell.Run "C:\Users\poh25\Videos\mini\C070.mp4"
   
   ElseIf Barcode = "C071" Then
       shell.Run "C:\Users\poh25\Videos\mini\C071.mp4"
   
   ElseIf Barcode = "C072" Then
       shell.Run "C:\Users\poh25\Videos\mini\C072.mp4"
   
   ElseIf Barcode = "C073" Then
       shell.Run "C:\Users\poh25\Videos\mini\C073.mp4"
   
   ElseIf Barcode = "C074" Then
       shell.Run "C:\Users\poh25\Videos\mini\C074.mp4"
   
   ElseIf Barcode = "C075" Then
       shell.Run "C:\Users\poh25\Videos\mini\C075.mp4"
   
   ElseIf Barcode = "C076" Then
       shell.Run "C:\Users\poh25\Videos\mini\C076.mp4"
   
   ElseIf Barcode = "C077" Then
       shell.Run "C:\Users\poh25\Videos\mini\C077.mp4"
   
   ElseIf Barcode = "C078" Then
       shell.Run "C:\Users\poh25\Videos\mini\C078.mp4"
   
   ElseIf Barcode = "C079" Then
       shell.Run "C:\Users\poh25\Videos\mini\C079.mp4"
   
   ElseIf Barcode = "C080" Then
       shell.Run "C:\Users\poh25\Videos\mini\C080.mp4"
   
   ElseIf Barcode = "C081" Then
       shell.Run "C:\Users\poh25\Videos\mini\C081.mp4"
   
   ElseIf Barcode = "C082" Then
       shell.Run "C:\Users\poh25\Videos\mini\C082.mp4"
   
   ElseIf Barcode = "C083" Then
       shell.Run "C:\Users\poh25\Videos\mini\C083.mp4"
   
   ElseIf Barcode = "C084" Then
       shell.Run "C:\Users\poh25\Videos\mini\C084.mp4"
   
   ElseIf Barcode = "C085" Then
       shell.Run "C:\Users\poh25\Videos\mini\C085.mp4"
   
   ElseIf Barcode = "C086" Then
       shell.Run "C:\Users\poh25\Videos\mini\C086.mp4"
   
   ElseIf Barcode = "C087" Then
       shell.Run "C:\Users\poh25\Videos\mini\C087.mp4"
   
   ElseIf Barcode = "C088" Then
       shell.Run "C:\Users\poh25\Videos\mini\C088.mp4"
   
   ElseIf Barcode = "C089" Then
       shell.Run "C:\Users\poh25\Videos\mini\C089.mp4"
   
   ElseIf Barcode = "C090" Then
       shell.Run "C:\Users\poh25\Videos\mini\C090.mp4"
   
   ElseIf Barcode = "C091" Then
       shell.Run "C:\Users\poh25\Videos\mini\C091.mp4"
   
   ElseIf Barcode = "C092" Then
       shell.Run "C:\Users\poh25\Videos\mini\C092.mp4"
   
   ElseIf Barcode = "C093" Then
       shell.Run "C:\Users\poh25\Videos\mini\C093.mp4"
   
   ElseIf Barcode = "C094" Then
       shell.Run "C:\Users\poh25\Videos\mini\C094.mp4"
   
   ElseIf Barcode = "C095" Then
       shell.Run "C:\Users\poh25\Videos\mini\C095.mp4"
   
   ElseIf Barcode = "C096" Then
       shell.Run "C:\Users\poh25\Videos\mini\C096.mp4"
   
   ElseIf Barcode = "C097" Then
       shell.Run "C:\Users\poh25\Videos\mini\C097.mp4"
   
   ElseIf Barcode = "C098" Then
       shell.Run "C:\Users\poh25\Videos\mini\C098.mp4"
   
   ElseIf Barcode = "C099" Then
       shell.Run "C:\Users\poh25\Videos\mini\C099.mp4"
   
   ElseIf Barcode = "C100" Then
       shell.Run "C:\Users\poh25\Videos\mini\C100.mp4"
   
   ElseIf Barcode = "D001" Then
       shell.Run "C:\Users\poh25\Videos\mini\D001.mp4"
   
   ElseIf Barcode = "D002" Then
       shell.Run "C:\Users\poh25\Videos\mini\D002.mp4"
   
   ElseIf Barcode = "D003" Then
       shell.Run "C:\Users\poh25\Videos\mini\D003.mp4"
   
   ElseIf Barcode = "D004" Then
       shell.Run "C:\Users\poh25\Videos\mini\D004.mp4"
   
   ElseIf Barcode = "D005" Then
       shell.Run "C:\Users\poh25\Videos\mini\D005.mp4"
   
   ElseIf Barcode = "D006" Then
       shell.Run "C:\Users\poh25\Videos\mini\D006.mp4"
   
   ElseIf Barcode = "D007" Then
       shell.Run "C:\Users\poh25\Videos\mini\D007.mp4"
   
   ElseIf Barcode = "D008" Then
       shell.Run "C:\Users\poh25\Videos\mini\D008.mp4"
   
   ElseIf Barcode = "D009" Then
       shell.Run "C:\Users\poh25\Videos\mini\D009.mp4"
   
   ElseIf Barcode = "D010" Then
       shell.Run "C:\Users\poh25\Videos\mini\D010.mp4"
   
   ElseIf Barcode = "D011" Then
       shell.Run "C:\Users\poh25\Videos\mini\D011.mp4"
   
   ElseIf Barcode = "D012" Then
       shell.Run "C:\Users\poh25\Videos\mini\D012.mp4"
   
   ElseIf Barcode = "D013" Then
       shell.Run "C:\Users\poh25\Videos\mini\D013.mp4"
   
   ElseIf Barcode = "D014" Then
       shell.Run "C:\Users\poh25\Videos\mini\D014.mp4"
   
   ElseIf Barcode = "D015" Then
       shell.Run "C:\Users\poh25\Videos\mini\D015.mp4"
   
   ElseIf Barcode = "D016" Then
       shell.Run "C:\Users\poh25\Videos\mini\D016.mp4"
   
   ElseIf Barcode = "D017" Then
       shell.Run "C:\Users\poh25\Videos\mini\D017.mp4"
   
   ElseIf Barcode = "D018" Then
       shell.Run "C:\Users\poh25\Videos\mini\D018.mp4"
   
   ElseIf Barcode = "D019" Then
       shell.Run "C:\Users\poh25\Videos\mini\D019.mp4"
   
   ElseIf Barcode = "D020" Then
       shell.Run "C:\Users\poh25\Videos\mini\D020.mp4"
   
   ElseIf Barcode = "D021" Then
       shell.Run "C:\Users\poh25\Videos\mini\D021.mp4"
   
   ElseIf Barcode = "D022" Then
       shell.Run "C:\Users\poh25\Videos\mini\D022.mp4"
   
   ElseIf Barcode = "D023" Then
       shell.Run "C:\Users\poh25\Videos\mini\D023.mp4"
   
   ElseIf Barcode = "D024" Then
       shell.Run "C:\Users\poh25\Videos\mini\D024.mp4"
   
   ElseIf Barcode = "D025" Then
       shell.Run "C:\Users\poh25\Videos\mini\D025.mp4"
   
   ElseIf Barcode = "D026" Then
       shell.Run "C:\Users\poh25\Videos\mini\D026.mp4"
   
   ElseIf Barcode = "D027" Then
       shell.Run "C:\Users\poh25\Videos\mini\D027.mp4"
   
   ElseIf Barcode = "D028" Then
       shell.Run "C:\Users\poh25\Videos\mini\D028.mp4"
   
   ElseIf Barcode = "D029" Then
       shell.Run "C:\Users\poh25\Videos\mini\D029.mp4"
   
   ElseIf Barcode = "D030" Then
       shell.Run "C:\Users\poh25\Videos\mini\D030.mp4"
   
   ElseIf Barcode = "D031" Then
       shell.Run "C:\Users\poh25\Videos\mini\D031.mp4"
   
   ElseIf Barcode = "D032" Then
       shell.Run "C:\Users\poh25\Videos\mini\D032.mp4"
   
   ElseIf Barcode = "D033" Then
       shell.Run "C:\Users\poh25\Videos\mini\D033.mp4"
   
   ElseIf Barcode = "D034" Then
       shell.Run "C:\Users\poh25\Videos\mini\D034.mp4"
   
   ElseIf Barcode = "D035" Then
       shell.Run "C:\Users\poh25\Videos\mini\D035.mp4"
   
   ElseIf Barcode = "D036" Then
       shell.Run "C:\Users\poh25\Videos\mini\D036.mp4"
   
   ElseIf Barcode = "D037" Then
       shell.Run "C:\Users\poh25\Videos\mini\D037.mp4"
   
   ElseIf Barcode = "D038" Then
       shell.Run "C:\Users\poh25\Videos\mini\D038.mp4"
   
   ElseIf Barcode = "D039" Then
       shell.Run "C:\Users\poh25\Videos\mini\D039.mp4"
   
   ElseIf Barcode = "D040" Then
       shell.Run "C:\Users\poh25\Videos\mini\D040.mp4"
   
   ElseIf Barcode = "D041" Then
       shell.Run "C:\Users\poh25\Videos\mini\D041.mp4"
   
   ElseIf Barcode = "D042" Then
       shell.Run "C:\Users\poh25\Videos\mini\D042.mp4"
   
   ElseIf Barcode = "D043" Then
       shell.Run "C:\Users\poh25\Videos\mini\D043.mp4"
   
   ElseIf Barcode = "D044" Then
       shell.Run "C:\Users\poh25\Videos\mini\D044.mp4"
   
   ElseIf Barcode = "D045" Then
       shell.Run "C:\Users\poh25\Videos\mini\D045.mp4"
   
   ElseIf Barcode = "D046" Then
       shell.Run "C:\Users\poh25\Videos\mini\D046.mp4"
   
   ElseIf Barcode = "D047" Then
       shell.Run "C:\Users\poh25\Videos\mini\D047.mp4"
   
   ElseIf Barcode = "D048" Then
       shell.Run "C:\Users\poh25\Videos\mini\D048.mp4"
   
   ElseIf Barcode = "D049" Then
       shell.Run "C:\Users\poh25\Videos\mini\D049.mp4"
   
   ElseIf Barcode = "D050" Then
       shell.Run "C:\Users\poh25\Videos\mini\D050.mp4"
   
   ElseIf Barcode = "D051" Then
       shell.Run "C:\Users\poh25\Videos\mini\D051.mp4"
   
   ElseIf Barcode = "D052" Then
       shell.Run "C:\Users\poh25\Videos\mini\D052.mp4"
   
   ElseIf Barcode = "D053" Then
       shell.Run "C:\Users\poh25\Videos\mini\D053.mp4"
   
   ElseIf Barcode = "D054" Then
       shell.Run "C:\Users\poh25\Videos\mini\D054.mp4"
   
   ElseIf Barcode = "D055" Then
       shell.Run "C:\Users\poh25\Videos\mini\D055.mp4"
   
   ElseIf Barcode = "D056" Then
       shell.Run "C:\Users\poh25\Videos\mini\D056.mp4"
   
   ElseIf Barcode = "D057" Then
       shell.Run "C:\Users\poh25\Videos\mini\D057.mp4"
   
   ElseIf Barcode = "D058" Then
       shell.Run "C:\Users\poh25\Videos\mini\D058.mp4"
   
   ElseIf Barcode = "D059" Then
       shell.Run "C:\Users\poh25\Videos\mini\D059.mp4"
   
   ElseIf Barcode = "D060" Then
       shell.Run "C:\Users\poh25\Videos\mini\D060.mp4"
   
   ElseIf Barcode = "D061" Then
       shell.Run "C:\Users\poh25\Videos\mini\D061.mp4"
   
   ElseIf Barcode = "D062" Then
       shell.Run "C:\Users\poh25\Videos\mini\D062.mp4"
   
   ElseIf Barcode = "D063" Then
       shell.Run "C:\Users\poh25\Videos\mini\D063.mp4"
   
   ElseIf Barcode = "D064" Then
       shell.Run "C:\Users\poh25\Videos\mini\D064.mp4"
   
   ElseIf Barcode = "D065" Then
       shell.Run "C:\Users\poh25\Videos\mini\D065.mp4"
   
   ElseIf Barcode = "D066" Then
       shell.Run "C:\Users\poh25\Videos\mini\D066.mp4"
   
   ElseIf Barcode = "D067" Then
       shell.Run "C:\Users\poh25\Videos\mini\D067.mp4"
   
   ElseIf Barcode = "D068" Then
       shell.Run "C:\Users\poh25\Videos\mini\D068.mp4"
   
   ElseIf Barcode = "D069" Then
       shell.Run "C:\Users\poh25\Videos\mini\D069.mp4"
   
   ElseIf Barcode = "D070" Then
       shell.Run "C:\Users\poh25\Videos\mini\D070.mp4"
   
   ElseIf Barcode = "D071" Then
       shell.Run "C:\Users\poh25\Videos\mini\D071.mp4"
   
   ElseIf Barcode = "D072" Then
       shell.Run "C:\Users\poh25\Videos\mini\D072.mp4"
   
   ElseIf Barcode = "D073" Then
       shell.Run "C:\Users\poh25\Videos\mini\D073.mp4"
   
   ElseIf Barcode = "D074" Then
       shell.Run "C:\Users\poh25\Videos\mini\D074.mp4"
   
   ElseIf Barcode = "D075" Then
       shell.Run "C:\Users\poh25\Videos\mini\D075.mp4"
   
   ElseIf Barcode = "D076" Then
       shell.Run "C:\Users\poh25\Videos\mini\D076.mp4"
   
   ElseIf Barcode = "D077" Then
       shell.Run "C:\Users\poh25\Videos\mini\D077.mp4"
   
   ElseIf Barcode = "D078" Then
       shell.Run "C:\Users\poh25\Videos\mini\D078.mp4"
   
   ElseIf Barcode = "D079" Then
       shell.Run "C:\Users\poh25\Videos\mini\D079.mp4"
   
   ElseIf Barcode = "D080" Then
       shell.Run "C:\Users\poh25\Videos\mini\D080.mp4"
   
   ElseIf Barcode = "D081" Then
       shell.Run "C:\Users\poh25\Videos\mini\D081.mp4"
   
   ElseIf Barcode = "D082" Then
       shell.Run "C:\Users\poh25\Videos\mini\D082.mp4"
   
   ElseIf Barcode = "D083" Then
       shell.Run "C:\Users\poh25\Videos\mini\D083.mp4"
   
